(* IEC 61131-3 sources: deprecated-refusr-repo/samples (part 19) *)

(* ---- RND-EXPR_audio-kudos-nifty.st ---- *)
(*
This code implements a randomly grown symbolic expression:

IN3 | (xor(xor(IN43 | ((xor(xor(!(((xor(xor(IN13, IN9 | false), xor(xor(IN25, IN14), IN11))) | (xor(xor(xor(xor(IN36, IN12), IN39), IN13 & IN34), IN47))) | (xor(xor(IN5, (IN1 & IN27) | (!(IN46))), !(!(IN21))))), IN37), xor(xor(!(!(IN1)), !((xor(xor(IN30, false), xor(xor(IN49, IN30), IN25))) & (!(xor(xor(IN21, IN32), IN27))))), (xor(xor(!(xor(xor(IN12, IN39), IN41)), (IN22 & IN36) & (IN27 | IN16)), IN15)) | (!((IN24 | IN40) | (!(IN45))))))) & (xor(xor(!((!((false | IN41) & (!(IN49)))) | (((IN6 & IN32) & IN14) & (!(IN27 & IN33)))), xor(xor(xor(xor(IN38, (!(IN43 & IN26)) & ((IN34 & IN40) & (IN5 & IN12))), !(xor(xor(xor(xor(IN8, IN19), IN14), IN15 & IN11), IN30 & IN31))), ((xor(xor(IN24, IN1 | IN19), true | IN1)) & IN27) & ((IN25 | (IN21 | IN15)) & (IN13 & (IN19 & IN30)))), (((IN33 & true) | (IN35 | IN7)) & (xor(xor(true | IN16, IN48), IN43 & IN22))) & ((!(xor(xor(IN38, IN35), IN42))) & (!(IN39))))), xor(xor(IN6, (xor(xor(xor(xor(xor(xor(IN6, IN45), IN26), !(IN35)), IN32 | IN15), (!(IN15)) & (IN36 | IN34)), (xor(xor(IN47, IN47), IN44)) & (!(IN14)))) & (((IN13 & IN4) | (IN1 | IN38)) | ((IN46 & IN11) & (IN32 | IN24)))), IN18)))), !(xor(xor(!(!(xor(xor(IN1, !((xor(xor(IN33, IN25), IN4)) & (IN40 | IN38))), xor(xor(IN12, xor(xor(xor(xor(IN24, IN3), IN41), !(IN13)), IN50 & IN19)), (xor(xor(IN37, IN25), IN21)) | IN4)))), !(IN23)), (!((!((!(IN20)) & (IN23 & IN14))) | (IN43 | (xor(xor(IN27 & IN10, IN34), xor(xor(IN31, IN6), IN4)))))) | ((((!(IN27 | IN41)) | ((IN12 | IN28) | IN22)) & IN29) & (IN50 & (IN1 | ((xor(xor(IN49, IN28), IN4)) | (IN33 & IN4)))))))), (!((xor(xor((!(xor(xor(!(IN27), xor(xor(IN4, IN6), IN33)), IN31 & true))) | (!((xor(xor(IN40, IN39), IN27)) & (IN13 & IN12))), (((IN25 & IN4) & (!(IN17))) & (xor(xor(true | IN33, IN38), IN16))) & (xor(xor(IN44, !(xor(xor(IN27, IN40), IN11))), xor(xor(IN36 & IN37, IN15 | IN33), IN21)))), IN17 | (IN33 | ((IN2 & IN1) | IN33)))) & (((((IN33 & false) | (IN37 | IN18)) | (!(IN28))) & (xor(xor((IN38 | IN8) | (!(IN12)), !(IN1 | IN1)), IN30))) | (xor(xor((xor(xor(IN47 & IN24, IN47 & IN36), IN9)) & (!(IN31 & IN18)), xor(xor((!(IN49)) & IN4, (IN44 & IN19) | (IN26 | IN18)), !(!(IN34)))), !(IN32 & (IN33 | IN47))))))) | ((xor(xor(IN13, (!(true | (xor(xor(!(IN35), IN15 | IN4), xor(xor(IN35, IN27), IN15))))) & ((xor(xor(!(IN18 & IN31), IN22 | (IN7 & IN11)), !(xor(xor(IN37, IN45), IN24)))) & IN23)), IN35)) & IN5)))

*)

FUNCTION_BLOCK F_CollectInput
  VAR_IN_OUT
      Data : ARRAY[1..50] OF BOOL;
  END_VAR
  VAR_INPUT
      TICK  : BOOL := 0;
      IN1   : BOOL := 0;
      IN2   : BOOL := 0;
      IN3   : BOOL := 0;
      IN4   : BOOL := 0;
      IN5   : BOOL := 0;
      RESET : BOOL := FALSE;
  END_VAR
  VAR_OUTPUT
      Finished : BOOL;
  END_VAR
  VAR
      j    : USINT := 1;
      tock : BOOL  := 0;
  END_VAR
  IF NOT RESET AND tock = NOT TICK THEN
      Data[j]   := IN1;
      Data[j+1] := IN2;
      Data[j+2] := IN3;
      Data[j+3] := IN4;
      Data[j+4] := IN5;
      j := j + 5;
      tock := TICK;
  ELSE
      j := 1;
      tock := 0;
  END_IF;
  Finished := (j > 50);
END_FUNCTION_BLOCK

PROGRAM Boiler
  VAR
    Data  : ARRAY[1..50] OF BOOL;
    Ready : BOOL;
    CollectInput : F_CollectInput;
  END_VAR
  VAR
    TICK     AT %IX1.0 : BOOL;
    IN1      AT %IX0.3 : BOOL;
    IN2      AT %IX0.4 : BOOL;
    IN3      AT %IX0.5 : BOOL;
    IN4      AT %IX0.6 : BOOL;
    IN5      AT %IX0.7 : BOOL;
    OutReady AT %QX0.0 : BOOL := FALSE;
    FeedNext AT %QX0.1 : BOOL := FALSE;
    Out      AT %QX0.2 : BOOL;
  END_VAR
  CollectInput(TICK:=TICK, IN1:=IN1, IN2:=IN2, IN3:=IN3, IN4:=IN4, IN5:=IN5);
  Ready := CollectInput.Finished;
  FeedNext := 1;
  IF Ready THEN
    Out := (Data[3] OR (((Data[43] OR ((((NOT ((((Data[13] XOR (Data[9] OR FALSE)) XOR ((Data[25] XOR Data[14]) XOR Data[11])) OR ((((Data[36] XOR Data[12]) XOR Data[39]) XOR (Data[13] AND Data[34])) XOR Data[47])) OR ((Data[5] XOR ((Data[1] AND Data[27]) OR (NOT Data[46]))) XOR (NOT (NOT Data[21]))))) XOR Data[37]) XOR (((NOT (NOT Data[1])) XOR (NOT (((Data[30] XOR FALSE) XOR ((Data[49] XOR Data[30]) XOR Data[25])) AND (NOT ((Data[21] XOR Data[32]) XOR Data[27]))))) XOR ((((NOT ((Data[12] XOR Data[39]) XOR Data[41])) XOR ((Data[22] AND Data[36]) AND (Data[27] OR Data[16]))) XOR Data[15]) OR (NOT ((Data[24] OR Data[40]) OR (NOT Data[45])))))) AND (((NOT ((NOT ((FALSE OR Data[41]) AND (NOT Data[49]))) OR (((Data[6] AND Data[32]) AND Data[14]) AND (NOT (Data[27] AND Data[33]))))) XOR ((((Data[38] XOR ((NOT (Data[43] AND Data[26])) AND ((Data[34] AND Data[40]) AND (Data[5] AND Data[12])))) XOR (NOT ((((Data[8] XOR Data[19]) XOR Data[14]) XOR (Data[15] AND Data[11])) XOR (Data[30] AND Data[31])))) XOR ((((Data[24] XOR (Data[1] OR Data[19])) XOR (TRUE OR Data[1])) AND Data[27]) AND ((Data[25] OR (Data[21] OR Data[15])) AND (Data[13] AND (Data[19] AND Data[30]))))) XOR ((((Data[33] AND TRUE) OR (Data[35] OR Data[7])) AND (((TRUE OR Data[16]) XOR Data[48]) XOR (Data[43] AND Data[22]))) AND ((NOT ((Data[38] XOR Data[35]) XOR Data[42])) AND (NOT Data[39]))))) XOR ((Data[6] XOR (((((((Data[6] XOR Data[45]) XOR Data[26]) XOR (NOT Data[35])) XOR (Data[32] OR Data[15])) XOR ((NOT Data[15]) AND (Data[36] OR Data[34]))) XOR (((Data[47] XOR Data[47]) XOR Data[44]) AND (NOT Data[14]))) AND (((Data[13] AND Data[4]) OR (Data[1] OR Data[38])) OR ((Data[46] AND Data[11]) AND (Data[32] OR Data[24]))))) XOR Data[18])))) XOR (NOT (((NOT (NOT ((Data[1] XOR (NOT (((Data[33] XOR Data[25]) XOR Data[4]) AND (Data[40] OR Data[38])))) XOR ((Data[12] XOR ((((Data[24] XOR Data[3]) XOR Data[41]) XOR (NOT Data[13])) XOR (Data[50] AND Data[19]))) XOR (((Data[37] XOR Data[25]) XOR Data[21]) OR Data[4]))))) XOR (NOT Data[23])) XOR ((NOT ((NOT ((NOT Data[20]) AND (Data[23] AND Data[14]))) OR (Data[43] OR (((Data[27] AND Data[10]) XOR Data[34]) XOR ((Data[31] XOR Data[6]) XOR Data[4]))))) OR ((((NOT (Data[27] OR Data[41])) OR ((Data[12] OR Data[28]) OR Data[22])) AND Data[29]) AND (Data[50] AND (Data[1] OR (((Data[49] XOR Data[28]) XOR Data[4]) OR (Data[33] AND Data[4]))))))))) XOR ((NOT (((((NOT (((NOT Data[27]) XOR ((Data[4] XOR Data[6]) XOR Data[33])) XOR (Data[31] AND TRUE))) OR (NOT (((Data[40] XOR Data[39]) XOR Data[27]) AND (Data[13] AND Data[12])))) XOR ((((Data[25] AND Data[4]) AND (NOT Data[17])) AND (((TRUE OR Data[33]) XOR Data[38]) XOR Data[16])) AND ((Data[44] XOR (NOT ((Data[27] XOR Data[40]) XOR Data[11]))) XOR (((Data[36] AND Data[37]) XOR (Data[15] OR Data[33])) XOR Data[21])))) XOR (Data[17] OR (Data[33] OR ((Data[2] AND Data[1]) OR Data[33])))) AND (((((Data[33] AND FALSE) OR (Data[37] OR Data[18])) OR (NOT Data[28])) AND ((((Data[38] OR Data[8]) OR (NOT Data[12])) XOR (NOT (Data[1] OR Data[1]))) XOR Data[30])) OR ((((((Data[47] AND Data[24]) XOR (Data[47] AND Data[36])) XOR Data[9]) AND (NOT (Data[31] AND Data[18]))) XOR ((((NOT Data[49]) AND Data[4]) XOR ((Data[44] AND Data[19]) OR (Data[26] OR Data[18]))) XOR (NOT (NOT Data[34])))) XOR (NOT (Data[32] AND (Data[33] OR Data[47]))))))) OR (((Data[13] XOR ((NOT (TRUE OR (((NOT Data[35]) XOR (Data[15] OR Data[4])) XOR ((Data[35] XOR Data[27]) XOR Data[15])))) AND ((((NOT (Data[18] AND Data[31])) XOR (Data[22] OR (Data[7] AND Data[11]))) XOR (NOT ((Data[37] XOR Data[45]) XOR Data[24]))) AND Data[23]))) XOR Data[35]) AND Data[5]))));
    OutReady := 1;
    CollectInput(RESET:=TRUE);
  END_IF;
END_PROGRAM

CONFIGURATION Config0
  RESOURCE Res0 ON PLC
    TASK task0(INTERVAL := T#20ms,PRIORITY := 0);
    PROGRAM instance0 WITH task0 : Boiler;
  END_RESOURCE
END_CONFIGURATION

(* ---- RND-EXPR_awoke-fount-idled.st ---- *)
(*
This code implements a randomly grown symbolic expression:

!(xor(xor(IN7, (xor(xor(IN10 | (xor(xor(IN35 & (((xor(xor(IN23, IN37), IN21)) & (IN38 & IN15)) | (xor(xor(xor(xor(IN32, IN34), IN21), false & IN13), IN2 | IN26))), IN35 & (((xor(xor(IN7, IN2), false)) | (!(IN1))) | (xor(xor(!(IN25), xor(xor(IN45, IN1), IN42)), IN26 | IN16)))), xor(xor((xor(xor(!(IN35), IN47 | IN5), IN39 & IN10)) & ((xor(xor(IN16, IN37), IN23)) | (!(IN48))), !(IN46)), !(!(!(IN21)))))), IN28), false)) & (xor(xor(xor(xor((((xor(xor(xor(xor(IN46, IN37), IN44), IN29 & IN42), IN10 | false)) | (xor(xor(IN38 & false, IN30 & IN3), true))) | (((xor(xor(IN14, IN23), IN50)) & (xor(xor(IN24, IN27), IN22))) | ((xor(xor(IN18, IN21), IN34)) & (true | IN4)))) & (xor(xor((xor(xor(xor(xor(IN29, IN24), true), IN12 & IN14), IN2 | IN19)) & (!(IN30 & IN14)), (IN10 | (!(IN9))) | ((IN42 & IN44) & (IN33 & IN25))), IN5)), IN3 & ((xor(xor((IN36 & IN29) & (IN6 | IN45), xor(xor(!(IN2), !(IN10)), IN20)), IN43)) & (!((IN33 | IN35) | (xor(xor(IN50, IN35), IN48)))))), xor(xor((xor(xor(!(!(IN46)), IN34 | (IN35 | IN49)), (!(IN34)) & (IN10 & IN4))) & (IN15 | IN25), IN22), (xor(xor(xor(xor(IN30, IN12 | IN23), !(IN14)), IN1), (IN4 | IN32) & (!(IN48)))) | (((xor(xor(IN50, true), IN31)) & (xor(xor(IN22, IN32), IN34))) | (xor(xor(IN37, !(IN49)), IN22))))), xor(xor(!(xor(xor(xor(xor((IN48 & IN24) | (xor(xor(IN41, IN39), IN11)), IN14), IN11), IN39 & (!(IN10 | IN49))), IN44)), ((!(!(!(IN50)))) & ((xor(xor(IN35, !(IN50)), IN32 | IN49)) & (xor(xor(IN21 & IN42, true & IN25), IN4 & IN31)))) | (((!(IN21)) | (!(xor(xor(IN1, IN30), IN46)))) & (((IN6 | IN8) & (xor(xor(IN43, IN10), false))) | IN6))), xor(xor((xor(xor((IN34 | IN3) & (!(IN18)), (!(IN14)) & true), xor(xor(xor(xor(IN15, IN7), IN34), !(IN31)), IN20 | IN18))) | (((IN1 | IN1) & (IN5 | IN27)) | IN17), xor(xor((xor(xor(xor(xor(IN32, IN10), IN1), IN35 | IN32), IN8)) & (IN11 & (IN14 | IN16)), !((IN20 & IN44) | (IN6 | IN15))), (xor(xor(IN35 | IN40, !(IN35)), IN3 | IN48)) | (!(IN46)))), (!(IN14)) & IN7))), (xor(xor(!(xor(xor(IN18, xor(xor(IN24 & IN23, !(IN40)), xor(xor(IN27, IN31), IN35))), !(xor(xor(false, IN48), IN6)))), (!((IN23 | IN37) & (IN8 | IN41))) & IN25), IN5 | (((xor(xor(IN41, IN26), IN3)) & (IN46 | IN22)) | ((IN49 & IN45) & (IN42 & IN16))))) | ((((!(IN47)) | true) & (IN30 | ((IN46 & IN30) | (!(IN43))))) | (((xor(xor(IN37, !(IN40)), !(IN4))) | (IN11 & (!(IN40)))) | (xor(xor(xor(xor(IN46 | IN15, IN9 | IN2), !(IN15)), xor(xor(!(IN46), false), IN36 & IN44)), !(!(IN27))))))))), !(IN35 & (xor(xor((xor(xor(xor(xor(!(xor(xor(IN12, IN9), IN31)), (xor(xor(IN35, IN38), IN3)) | (xor(xor(IN47, IN13), IN8))), (IN36 & false) | (IN13 | IN46)), IN19), (IN47 & (IN46 | IN35)) | IN25)) & (xor(xor(xor(xor((IN14 | IN37) | (IN10 | IN3), IN39 & IN30), xor(xor(IN33 & IN5, xor(xor(IN39, IN48), IN16)), !(IN33))), !(IN38)), !(!(IN33 | IN3)))), IN48), IN20)))))

*)

FUNCTION_BLOCK F_CollectInput
  VAR_IN_OUT
      Data : ARRAY[1..50] OF BOOL;
  END_VAR
  VAR_INPUT
      TICK  : BOOL := 0;
      IN1   : BOOL := 0;
      IN2   : BOOL := 0;
      IN3   : BOOL := 0;
      IN4   : BOOL := 0;
      IN5   : BOOL := 0;
      RESET : BOOL := FALSE;
  END_VAR
  VAR_OUTPUT
      Finished : BOOL;
  END_VAR
  VAR
      j    : USINT := 1;
      tock : BOOL  := 0;
  END_VAR
  IF NOT RESET AND tock = NOT TICK THEN
      Data[j]   := IN1;
      Data[j+1] := IN2;
      Data[j+2] := IN3;
      Data[j+3] := IN4;
      Data[j+4] := IN5;
      j := j + 5;
      tock := TICK;
  ELSE
      j := 1;
      tock := 0;
  END_IF;
  Finished := (j > 50);
END_FUNCTION_BLOCK

PROGRAM Boiler
  VAR
    Data  : ARRAY[1..50] OF BOOL;
    Ready : BOOL;
    CollectInput : F_CollectInput;
  END_VAR
  VAR
    TICK     AT %IX1.0 : BOOL;
    IN1      AT %IX0.3 : BOOL;
    IN2      AT %IX0.4 : BOOL;
    IN3      AT %IX0.5 : BOOL;
    IN4      AT %IX0.6 : BOOL;
    IN5      AT %IX0.7 : BOOL;
    OutReady AT %QX0.0 : BOOL := FALSE;
    FeedNext AT %QX0.1 : BOOL := FALSE;
    Out      AT %QX0.2 : BOOL;
  END_VAR
  CollectInput(TICK:=TICK, IN1:=IN1, IN2:=IN2, IN3:=IN3, IN4:=IN4, IN5:=IN5);
  Ready := CollectInput.Finished;
  FeedNext := 1;
  IF Ready THEN
    Out := (NOT ((Data[7] XOR ((((Data[10] OR (((Data[35] AND ((((Data[23] XOR Data[37]) XOR Data[21]) AND (Data[38] AND Data[15])) OR ((((Data[32] XOR Data[34]) XOR Data[21]) XOR (FALSE AND Data[13])) XOR (Data[2] OR Data[26])))) XOR (Data[35] AND ((((Data[7] XOR Data[2]) XOR FALSE) OR (NOT Data[1])) OR (((NOT Data[25]) XOR ((Data[45] XOR Data[1]) XOR Data[42])) XOR (Data[26] OR Data[16]))))) XOR ((((((NOT Data[35]) XOR (Data[47] OR Data[5])) XOR (Data[39] AND Data[10])) AND (((Data[16] XOR Data[37]) XOR Data[23]) OR (NOT Data[48]))) XOR (NOT Data[46])) XOR (NOT (NOT (NOT Data[21])))))) XOR Data[28]) XOR FALSE) AND (((((((((((Data[46] XOR Data[37]) XOR Data[44]) XOR (Data[29] AND Data[42])) XOR (Data[10] OR FALSE)) OR (((Data[38] AND FALSE) XOR (Data[30] AND Data[3])) XOR TRUE)) OR ((((Data[14] XOR Data[23]) XOR Data[50]) AND ((Data[24] XOR Data[27]) XOR Data[22])) OR (((Data[18] XOR Data[21]) XOR Data[34]) AND (TRUE OR Data[4])))) AND (((((((Data[29] XOR Data[24]) XOR TRUE) XOR (Data[12] AND Data[14])) XOR (Data[2] OR Data[19])) AND (NOT (Data[30] AND Data[14]))) XOR ((Data[10] OR (NOT Data[9])) OR ((Data[42] AND Data[44]) AND (Data[33] AND Data[25])))) XOR Data[5])) XOR (Data[3] AND (((((Data[36] AND Data[29]) AND (Data[6] OR Data[45])) XOR (((NOT Data[2]) XOR (NOT Data[10])) XOR Data[20])) XOR Data[43]) AND (NOT ((Data[33] OR Data[35]) OR ((Data[50] XOR Data[35]) XOR Data[48])))))) XOR ((((((NOT (NOT Data[46])) XOR (Data[34] OR (Data[35] OR Data[49]))) XOR ((NOT Data[34]) AND (Data[10] AND Data[4]))) AND (Data[15] OR Data[25])) XOR Data[22]) XOR (((((Data[30] XOR (Data[12] OR Data[23])) XOR (NOT Data[14])) XOR Data[1]) XOR ((Data[4] OR Data[32]) AND (NOT Data[48]))) OR ((((Data[50] XOR TRUE) XOR Data[31]) AND ((Data[22] XOR Data[32]) XOR Data[34])) OR ((Data[37] XOR (NOT Data[49])) XOR Data[22]))))) XOR (((NOT ((((((Data[48] AND Data[24]) OR ((Data[41] XOR Data[39]) XOR Data[11])) XOR Data[14]) XOR Data[11]) XOR (Data[39] AND (NOT (Data[10] OR Data[49])))) XOR Data[44])) XOR (((NOT (NOT (NOT Data[50]))) AND (((Data[35] XOR (NOT Data[50])) XOR (Data[32] OR Data[49])) AND (((Data[21] AND Data[42]) XOR (TRUE AND Data[25])) XOR (Data[4] AND Data[31])))) OR (((NOT Data[21]) OR (NOT ((Data[1] XOR Data[30]) XOR Data[46]))) AND (((Data[6] OR Data[8]) AND ((Data[43] XOR Data[10]) XOR FALSE)) OR Data[6])))) XOR (((((((Data[34] OR Data[3]) AND (NOT Data[18])) XOR ((NOT Data[14]) AND TRUE)) XOR ((((Data[15] XOR Data[7]) XOR Data[34]) XOR (NOT Data[31])) XOR (Data[20] OR Data[18]))) OR (((Data[1] OR Data[1]) AND (Data[5] OR Data[27])) OR Data[17])) XOR (((((((Data[32] XOR Data[10]) XOR Data[1]) XOR (Data[35] OR Data[32])) XOR Data[8]) AND (Data[11] AND (Data[14] OR Data[16]))) XOR (NOT ((Data[20] AND Data[44]) OR (Data[6] OR Data[15])))) XOR ((((Data[35] OR Data[40]) XOR (NOT Data[35])) XOR (Data[3] OR Data[48])) OR (NOT Data[46])))) XOR ((NOT Data[14]) AND Data[7])))) XOR ((((NOT ((Data[18] XOR (((Data[24] AND Data[23]) XOR (NOT Data[40])) XOR ((Data[27] XOR Data[31]) XOR Data[35]))) XOR (NOT ((FALSE XOR Data[48]) XOR Data[6])))) XOR ((NOT ((Data[23] OR Data[37]) AND (Data[8] OR Data[41]))) AND Data[25])) XOR (Data[5] OR ((((Data[41] XOR Data[26]) XOR Data[3]) AND (Data[46] OR Data[22])) OR ((Data[49] AND Data[45]) AND (Data[42] AND Data[16]))))) OR ((((NOT Data[47]) OR TRUE) AND (Data[30] OR ((Data[46] AND Data[30]) OR (NOT Data[43])))) OR ((((Data[37] XOR (NOT Data[40])) XOR (NOT Data[4])) OR (Data[11] AND (NOT Data[40]))) OR (((((Data[46] OR Data[15]) XOR (Data[9] OR Data[2])) XOR (NOT Data[15])) XOR (((NOT Data[46]) XOR FALSE) XOR (Data[36] AND Data[44]))) XOR (NOT (NOT Data[27]))))))))) XOR (NOT (Data[35] AND ((((((((NOT ((Data[12] XOR Data[9]) XOR Data[31])) XOR (((Data[35] XOR Data[38]) XOR Data[3]) OR ((Data[47] XOR Data[13]) XOR Data[8]))) XOR ((Data[36] AND FALSE) OR (Data[13] OR Data[46]))) XOR Data[19]) XOR ((Data[47] AND (Data[46] OR Data[35])) OR Data[25])) AND ((((((Data[14] OR Data[37]) OR (Data[10] OR Data[3])) XOR (Data[39] AND Data[30])) XOR (((Data[33] AND Data[5]) XOR ((Data[39] XOR Data[48]) XOR Data[16])) XOR (NOT Data[33]))) XOR (NOT Data[38])) XOR (NOT (NOT (Data[33] OR Data[3]))))) XOR Data[48]) XOR Data[20])))));
    OutReady := 1;
    CollectInput(RESET:=TRUE);
  END_IF;
END_PROGRAM

CONFIGURATION Config0
  RESOURCE Res0 ON PLC
    TASK task0(INTERVAL := T#20ms,PRIORITY := 0);
    PROGRAM instance0 WITH task0 : Boiler;
  END_RESOURCE
END_CONFIGURATION

(* ---- RND-EXPR_balmy-flubs-lives.st ---- *)
(*
This code implements a randomly grown symbolic expression:

(!(IN49)) & IN46

*)

FUNCTION_BLOCK F_CollectInput
  VAR_IN_OUT
      Data : ARRAY[1..50] OF BOOL;
  END_VAR
  VAR_INPUT
      TICK  : BOOL := 0;
      IN1   : BOOL := 0;
      IN2   : BOOL := 0;
      IN3   : BOOL := 0;
      IN4   : BOOL := 0;
      IN5   : BOOL := 0;
      RESET : BOOL := FALSE;
  END_VAR
  VAR_OUTPUT
      Finished : BOOL;
  END_VAR
  VAR
      j    : USINT := 1;
      tock : BOOL  := 0;
  END_VAR
  IF NOT RESET AND tock = NOT TICK THEN
      Data[j]   := IN1;
      Data[j+1] := IN2;
      Data[j+2] := IN3;
      Data[j+3] := IN4;
      Data[j+4] := IN5;
      j := j + 5;
      tock := TICK;
  ELSE
      j := 1;
      tock := 0;
  END_IF;
  Finished := (j > 50);
END_FUNCTION_BLOCK

PROGRAM Boiler
  VAR
    Data  : ARRAY[1..50] OF BOOL;
    Ready : BOOL;
    CollectInput : F_CollectInput;
  END_VAR
  VAR
    TICK     AT %IX1.0 : BOOL;
    IN1      AT %IX0.3 : BOOL;
    IN2      AT %IX0.4 : BOOL;
    IN3      AT %IX0.5 : BOOL;
    IN4      AT %IX0.6 : BOOL;
    IN5      AT %IX0.7 : BOOL;
    OutReady AT %QX0.0 : BOOL := FALSE;
    FeedNext AT %QX0.1 : BOOL := FALSE;
    Out      AT %QX0.2 : BOOL;
  END_VAR
  CollectInput(TICK:=TICK, IN1:=IN1, IN2:=IN2, IN3:=IN3, IN4:=IN4, IN5:=IN5);
  Ready := CollectInput.Finished;
  FeedNext := 1;
  IF Ready THEN
    Out := ((NOT Data[49]) AND Data[46]);
    OutReady := 1;
    CollectInput(RESET:=TRUE);
  END_IF;
END_PROGRAM

CONFIGURATION Config0
  RESOURCE Res0 ON PLC
    TASK task0(INTERVAL := T#20ms,PRIORITY := 0);
    PROGRAM instance0 WITH task0 : Boiler;
  END_RESOURCE
END_CONFIGURATION

(* ---- RND-EXPR_baton-smear-tarot.st ---- *)
(*
This code implements a randomly grown symbolic expression:

xor(xor(!((((IN19 | ((!(xor(xor(IN42 | IN9, IN18), IN43))) & (IN45 & (!(xor(xor(IN20, IN7), IN15)))))) | (xor(xor(IN2, (((xor(xor(IN43, IN1), IN41)) | (xor(xor(IN13, IN45), IN31))) & ((IN14 & IN3) | (IN11 | IN19))) | IN16), IN5 | IN40))) & IN38) & (IN44 | (IN29 & IN45))), xor(xor(IN21, IN35 & (!(IN21))), (!(xor(xor(xor(xor((!(IN16 | (xor(xor(IN8, IN25), IN37)))) & IN21, IN12), (!((IN32 & IN11) & (IN26 | IN3))) | (xor(xor(xor(xor(IN18 | IN31, IN48 | IN23), IN26 & IN42), !(IN24)), (IN22 & IN13) & (IN25 | IN12)))), IN16), IN13))) | (((!((((IN13 & IN39) & (!(IN34))) | IN2) | (!(!(xor(xor(IN23, IN32), IN28)))))) | (xor(xor(xor(xor((xor(xor(IN38 & IN21, IN45 | IN35), IN21 & IN26)) | IN1, ((IN23 | IN23) | IN17) & (!(IN20 & IN9))), IN39), !(!(xor(xor(IN26 & IN43, IN40 & IN33), false | IN33)))), IN49))) | IN3))), (!(!(!(IN2 & IN26)))) & (xor(xor((xor(xor((xor(xor(IN27, xor(xor(IN42 & (!(IN35)), (IN3 | IN32) & (IN4 | IN35)), (!(IN32)) & IN47)), (xor(xor(xor(xor(IN13, IN2), IN28), IN9 | IN42), !(IN30))) | ((IN9 | IN14) & (IN44 & IN28)))) & (!(IN21 | ((IN1 | IN41) & (IN6 | IN3)))), !(((!(IN41)) | IN41) & (IN13 | ((IN13 & IN10) & (xor(xor(IN27, IN13), IN7)))))), !(xor(xor(IN18, IN9), (!(IN38 & IN26)) & (xor(xor(IN21 | IN41, xor(xor(IN23, IN37), IN28)), !(IN7))))))) & ((!(xor(xor((IN17 & (!(IN29))) & ((IN22 & IN31) | (xor(xor(IN13, IN47), IN2))), ((!(IN7)) | IN4) | (xor(xor(!(IN19), !(IN19)), IN31))), !((xor(xor(IN8, IN12), false)) & (IN25 | IN21))))) & (IN5 | (xor(xor(xor(xor(xor(xor(xor(xor(IN14, IN16), IN50), IN9), IN44), xor(xor(xor(xor(IN19, IN1), IN13), IN2 & IN36), IN40)), !(IN10 | IN39)), IN20), (IN4 & (!(IN21))) & (IN8 | (IN30 & IN12)))))), (xor(xor((!((xor(xor(IN50 | IN6, IN28 & IN9), IN23)) | (xor(xor(IN41 | IN44, IN7 | IN29), !(IN26))))) | (((xor(xor(IN4, IN43 | IN10), IN17 & IN40)) & ((IN49 & IN39) & (xor(xor(IN18, IN39), IN12)))) & (!(IN11 & (IN26 | IN30)))), IN13), IN2 | ((((xor(xor(IN32, IN41), IN4)) & IN43) & ((IN18 | IN10) | (xor(xor(IN22, IN16), IN42)))) & (IN22 | (xor(xor(IN18 & IN35, IN14), IN20 & IN8)))))) & (((xor(xor(((IN6 & IN44) | (xor(xor(IN11, IN45), true))) | IN11, true), xor(xor((xor(xor(IN8, true), IN25)) & (xor(xor(IN39, IN32), IN11)), !(IN21 | IN28)), IN6))) | ((xor(xor(IN14, (!(IN16)) & (!(IN29))), xor(xor(IN27 | IN23, IN13), xor(xor(IN12, IN25), IN31)))) | (xor(xor(xor(xor(IN11 | IN50, !(IN48)), !(IN48)), IN14), IN27)))) | (!(IN34 & (((IN3 | IN14) | (true & IN17)) & ((xor(xor(IN39, IN50), IN5)) | (IN4 | IN18))))))), IN5)))

*)

FUNCTION_BLOCK F_CollectInput
  VAR_IN_OUT
      Data : ARRAY[1..50] OF BOOL;
  END_VAR
  VAR_INPUT
      TICK  : BOOL := 0;
      IN1   : BOOL := 0;
      IN2   : BOOL := 0;
      IN3   : BOOL := 0;
      IN4   : BOOL := 0;
      IN5   : BOOL := 0;
      RESET : BOOL := FALSE;
  END_VAR
  VAR_OUTPUT
      Finished : BOOL;
  END_VAR
  VAR
      j    : USINT := 1;
      tock : BOOL  := 0;
  END_VAR
  IF NOT RESET AND tock = NOT TICK THEN
      Data[j]   := IN1;
      Data[j+1] := IN2;
      Data[j+2] := IN3;
      Data[j+3] := IN4;
      Data[j+4] := IN5;
      j := j + 5;
      tock := TICK;
  ELSE
      j := 1;
      tock := 0;
  END_IF;
  Finished := (j > 50);
END_FUNCTION_BLOCK

PROGRAM Boiler
  VAR
    Data  : ARRAY[1..50] OF BOOL;
    Ready : BOOL;
    CollectInput : F_CollectInput;
  END_VAR
  VAR
    TICK     AT %IX1.0 : BOOL;
    IN1      AT %IX0.3 : BOOL;
    IN2      AT %IX0.4 : BOOL;
    IN3      AT %IX0.5 : BOOL;
    IN4      AT %IX0.6 : BOOL;
    IN5      AT %IX0.7 : BOOL;
    OutReady AT %QX0.0 : BOOL := FALSE;
    FeedNext AT %QX0.1 : BOOL := FALSE;
    Out      AT %QX0.2 : BOOL;
  END_VAR
  CollectInput(TICK:=TICK, IN1:=IN1, IN2:=IN2, IN3:=IN3, IN4:=IN4, IN5:=IN5);
  Ready := CollectInput.Finished;
  FeedNext := 1;
  IF Ready THEN
    Out := (((NOT ((((Data[19] OR ((NOT (((Data[42] OR Data[9]) XOR Data[18]) XOR Data[43])) AND (Data[45] AND (NOT ((Data[20] XOR Data[7]) XOR Data[15]))))) OR ((Data[2] XOR (((((Data[43] XOR Data[1]) XOR Data[41]) OR ((Data[13] XOR Data[45]) XOR Data[31])) AND ((Data[14] AND Data[3]) OR (Data[11] OR Data[19]))) OR Data[16])) XOR (Data[5] OR Data[40]))) AND Data[38]) AND (Data[44] OR (Data[29] AND Data[45])))) XOR ((Data[21] XOR (Data[35] AND (NOT Data[21]))) XOR ((NOT ((((((NOT (Data[16] OR ((Data[8] XOR Data[25]) XOR Data[37]))) AND Data[21]) XOR Data[12]) XOR ((NOT ((Data[32] AND Data[11]) AND (Data[26] OR Data[3]))) OR (((((Data[18] OR Data[31]) XOR (Data[48] OR Data[23])) XOR (Data[26] AND Data[42])) XOR (NOT Data[24])) XOR ((Data[22] AND Data[13]) AND (Data[25] OR Data[12]))))) XOR Data[16]) XOR Data[13])) OR (((NOT ((((Data[13] AND Data[39]) AND (NOT Data[34])) OR Data[2]) OR (NOT (NOT ((Data[23] XOR Data[32]) XOR Data[28]))))) OR ((((((((Data[38] AND Data[21]) XOR (Data[45] OR Data[35])) XOR (Data[21] AND Data[26])) OR Data[1]) XOR (((Data[23] OR Data[23]) OR Data[17]) AND (NOT (Data[20] AND Data[9])))) XOR Data[39]) XOR (NOT (NOT (((Data[26] AND Data[43]) XOR (Data[40] AND Data[33])) XOR (FALSE OR Data[33]))))) XOR Data[49])) OR Data[3])))) XOR ((NOT (NOT (NOT (Data[2] AND Data[26])))) AND ((((((((Data[27] XOR (((Data[42] AND (NOT Data[35])) XOR ((Data[3] OR Data[32]) AND (Data[4] OR Data[35]))) XOR ((NOT Data[32]) AND Data[47]))) XOR (((((Data[13] XOR Data[2]) XOR Data[28]) XOR (Data[9] OR Data[42])) XOR (NOT Data[30])) OR ((Data[9] OR Data[14]) AND (Data[44] AND Data[28])))) AND (NOT (Data[21] OR ((Data[1] OR Data[41]) AND (Data[6] OR Data[3]))))) XOR (NOT (((NOT Data[41]) OR Data[41]) AND (Data[13] OR ((Data[13] AND Data[10]) AND ((Data[27] XOR Data[13]) XOR Data[7])))))) XOR (NOT ((Data[18] XOR Data[9]) XOR ((NOT (Data[38] AND Data[26])) AND (((Data[21] OR Data[41]) XOR ((Data[23] XOR Data[37]) XOR Data[28])) XOR (NOT Data[7])))))) AND ((NOT ((((Data[17] AND (NOT Data[29])) AND ((Data[22] AND Data[31]) OR ((Data[13] XOR Data[47]) XOR Data[2]))) XOR (((NOT Data[7]) OR Data[4]) OR (((NOT Data[19]) XOR (NOT Data[19])) XOR Data[31]))) XOR (NOT (((Data[8] XOR Data[12]) XOR FALSE) AND (Data[25] OR Data[21]))))) AND (Data[5] OR ((((((((Data[14] XOR Data[16]) XOR Data[50]) XOR Data[9]) XOR Data[44]) XOR ((((Data[19] XOR Data[1]) XOR Data[13]) XOR (Data[2] AND Data[36])) XOR Data[40])) XOR (NOT (Data[10] OR Data[39]))) XOR Data[20]) XOR ((Data[4] AND (NOT Data[21])) AND (Data[8] OR (Data[30] AND Data[12]))))))) XOR (((((NOT ((((Data[50] OR Data[6]) XOR (Data[28] AND Data[9])) XOR Data[23]) OR (((Data[41] OR Data[44]) XOR (Data[7] OR Data[29])) XOR (NOT Data[26])))) OR ((((Data[4] XOR (Data[43] OR Data[10])) XOR (Data[17] AND Data[40])) AND ((Data[49] AND Data[39]) AND ((Data[18] XOR Data[39]) XOR Data[12]))) AND (NOT (Data[11] AND (Data[26] OR Data[30]))))) XOR Data[13]) XOR (Data[2] OR (((((Data[32] XOR Data[41]) XOR Data[4]) AND Data[43]) AND ((Data[18] OR Data[10]) OR ((Data[22] XOR Data[16]) XOR Data[42]))) AND (Data[22] OR (((Data[18] AND Data[35]) XOR Data[14]) XOR (Data[20] AND Data[8])))))) AND (((((((Data[6] AND Data[44]) OR ((Data[11] XOR Data[45]) XOR TRUE)) OR Data[11]) XOR TRUE) XOR (((((Data[8] XOR TRUE) XOR Data[25]) AND ((Data[39] XOR Data[32]) XOR Data[11])) XOR (NOT (Data[21] OR Data[28]))) XOR Data[6])) OR (((Data[14] XOR ((NOT Data[16]) AND (NOT Data[29]))) XOR (((Data[27] OR Data[23]) XOR Data[13]) XOR ((Data[12] XOR Data[25]) XOR Data[31]))) OR (((((Data[11] OR Data[50]) XOR (NOT Data[48])) XOR (NOT Data[48])) XOR Data[14]) XOR Data[27]))) OR (NOT (Data[34] AND (((Data[3] OR Data[14]) OR (TRUE AND Data[17])) AND (((Data[39] XOR Data[50]) XOR Data[5]) OR (Data[4] OR Data[18])))))))) XOR Data[5])));
    OutReady := 1;
    CollectInput(RESET:=TRUE);
  END_IF;
END_PROGRAM

CONFIGURATION Config0
  RESOURCE Res0 ON PLC
    TASK task0(INTERVAL := T#20ms,PRIORITY := 0);
    PROGRAM instance0 WITH task0 : Boiler;
  END_RESOURCE
END_CONFIGURATION

(* ---- RND-EXPR_beads-fetal-heads.st ---- *)
(*
This code implements a randomly grown symbolic expression:

(((!((((!((IN5 & IN33) | (IN35 | IN14))) & (!(xor(xor(xor(xor(IN9, IN33), IN3), IN49 | IN12), IN43)))) & (IN16 | IN22)) | (IN9 | ((!(!(IN6 | IN26))) | (xor(xor(!(IN23 & true), (IN16 & IN22) | (!(IN20))), IN12)))))) | ((((xor(xor(xor(xor(IN28, (xor(xor(IN2, IN16), IN38)) & (xor(xor(IN24, IN21), IN24))), !(!(IN35))), !(IN31 & IN50)), xor(xor(xor(xor(!(IN26), xor(xor(IN1, IN45), IN39)), xor(xor(IN37, IN8), IN27)), xor(xor(IN1 | IN20, true & IN23), !(IN22))), xor(xor(!(IN39), xor(xor(IN1, IN47), IN27)), IN22 | IN16)))) | ((((!(IN26)) & (IN33 & IN22)) | ((xor(xor(IN45, IN43), IN41)) | (xor(xor(IN40, IN11), IN48)))) & ((xor(xor(IN24 | IN1, xor(xor(false, IN2), IN3)), IN5 | IN44)) | ((IN50 & IN2) | (!(IN49)))))) & (!(IN35))) | (xor(xor(!(!(!((IN50 | IN15) | (IN40 & IN2)))), ((((IN34 & IN30) | (IN45 | IN41)) & ((IN3 | IN38) | IN2)) & ((IN18 | (!(IN19))) | ((IN48 | IN30) & (!(IN7))))) | (!((xor(xor(IN29 | IN29, IN46 & IN22), IN18 | IN11)) & (!(IN49 & IN15))))), (!(xor(xor((!(IN26)) & IN35, (!(IN27)) & (IN23 | IN41)), IN49 | (!(IN47))))) & (!(!(xor(xor(xor(xor(IN8, IN50), IN23), xor(xor(IN6, IN18), IN22)), IN12 | IN7)))))))) & (xor(xor((((((!(xor(xor(IN14, IN6), IN3))) & IN4) | (!((IN14 & IN24) & (xor(xor(IN3, IN21), IN20))))) | ((((!(IN36)) & IN28) | IN2) & IN40)) | (!((IN13 | IN14) | (xor(xor((xor(xor(IN17, IN22), IN30)) & (IN35 | IN35), !(xor(xor(IN46, IN8), true))), !(IN22)))))) | (((!(IN50)) & (xor(xor(((xor(xor(IN26, IN26), IN31)) | (xor(xor(true, IN46), IN46))) | ((IN7 & IN17) & (xor(xor(IN5, IN38), IN21))), !((IN13 | IN22) & (IN16 | IN46))), xor(xor(xor(xor(IN37, IN36), xor(xor(IN2, IN44), IN18)), (IN28 & IN19) & (IN37 | IN20)), (IN24 & IN34) & (IN43 & IN45))))) | (IN39 | (((!(IN12)) | (IN21 | (!(IN38)))) & ((xor(xor(!(IN28), IN35 & IN29), !(IN50))) & ((xor(xor(IN42, IN19), IN47)) | IN42))))), xor(xor(!(xor(xor((((IN45 & IN48) & (xor(xor(IN21, IN32), IN36))) | ((IN20 | IN25) | (!(IN44)))) | (((!(IN28)) & IN15) | ((!(IN43)) | IN44)), xor(xor(xor(xor(IN7 | (xor(xor(IN43, IN3), IN10)), (!(IN1)) & IN48), !(xor(xor(IN34, IN19), IN42))), xor(xor((!(IN46)) | (IN32 & IN3), xor(xor(IN6 | IN20, !(IN29)), false & IN14)), !(!(IN20)))), xor(xor((xor(xor(IN24, IN27), IN37)) & IN26, !(IN33 & IN46)), !(xor(xor(IN7, IN41), IN38))))), xor(xor(!(!(IN26)), IN50), ((IN28 & IN17) & (xor(xor(IN4, IN38), IN9))) | ((IN16 | IN31) & (!(IN32)))))), !((!(!(!(xor(xor(IN9, IN1), IN39))))) & (!(IN1 & (!(xor(xor(IN20, IN38), false))))))), IN17)), xor(xor(xor(xor(((!(IN16 & (IN49 & IN24))) | (xor(xor((xor(xor(IN27, IN22), IN3)) | (xor(xor(false, IN46), IN40)), !(xor(xor(IN42, IN4), IN32))), IN22 & (xor(xor(IN8, IN30), IN3))))) | ((xor(xor(IN27 | (IN38 & IN36), xor(xor(IN24 | IN12, IN1 & IN37), !(IN39))), !(IN50 & IN47))) & (!((xor(xor(IN16, IN8), IN26)) | (IN49 | IN40)))), xor(xor(!(xor(xor(true, xor(xor(true, IN47), IN5 & IN29)), xor(xor(IN7 & IN8, IN19), !(IN23)))), (!(!(!(IN6)))) & IN9), true)), IN29), IN48), IN2)))) | IN11

*)

FUNCTION_BLOCK F_CollectInput
  VAR_IN_OUT
      Data : ARRAY[1..50] OF BOOL;
  END_VAR
  VAR_INPUT
      TICK  : BOOL := 0;
      IN1   : BOOL := 0;
      IN2   : BOOL := 0;
      IN3   : BOOL := 0;
      IN4   : BOOL := 0;
      IN5   : BOOL := 0;
      RESET : BOOL := FALSE;
  END_VAR
  VAR_OUTPUT
      Finished : BOOL;
  END_VAR
  VAR
      j    : USINT := 1;
      tock : BOOL  := 0;
  END_VAR
  IF NOT RESET AND tock = NOT TICK THEN
      Data[j]   := IN1;
      Data[j+1] := IN2;
      Data[j+2] := IN3;
      Data[j+3] := IN4;
      Data[j+4] := IN5;
      j := j + 5;
      tock := TICK;
  ELSE
      j := 1;
      tock := 0;
  END_IF;
  Finished := (j > 50);
END_FUNCTION_BLOCK

PROGRAM Boiler
  VAR
    Data  : ARRAY[1..50] OF BOOL;
    Ready : BOOL;
    CollectInput : F_CollectInput;
  END_VAR
  VAR
    TICK     AT %IX1.0 : BOOL;
    IN1      AT %IX0.3 : BOOL;
    IN2      AT %IX0.4 : BOOL;
    IN3      AT %IX0.5 : BOOL;
    IN4      AT %IX0.6 : BOOL;
    IN5      AT %IX0.7 : BOOL;
    OutReady AT %QX0.0 : BOOL := FALSE;
    FeedNext AT %QX0.1 : BOOL := FALSE;
    Out      AT %QX0.2 : BOOL;
  END_VAR
  CollectInput(TICK:=TICK, IN1:=IN1, IN2:=IN2, IN3:=IN3, IN4:=IN4, IN5:=IN5);
  Ready := CollectInput.Finished;
  FeedNext := 1;
  IF Ready THEN
    Out := ((((NOT ((((NOT ((Data[5] AND Data[33]) OR (Data[35] OR Data[14]))) AND (NOT ((((Data[9] XOR Data[33]) XOR Data[3]) XOR (Data[49] OR Data[12])) XOR Data[43]))) AND (Data[16] OR Data[22])) OR (Data[9] OR ((NOT (NOT (Data[6] OR Data[26]))) OR (((NOT (Data[23] AND TRUE)) XOR ((Data[16] AND Data[22]) OR (NOT Data[20]))) XOR Data[12]))))) OR (((((((Data[28] XOR (((Data[2] XOR Data[16]) XOR Data[38]) AND ((Data[24] XOR Data[21]) XOR Data[24]))) XOR (NOT (NOT Data[35]))) XOR (NOT (Data[31] AND Data[50]))) XOR (((((NOT Data[26]) XOR ((Data[1] XOR Data[45]) XOR Data[39])) XOR ((Data[37] XOR Data[8]) XOR Data[27])) XOR (((Data[1] OR Data[20]) XOR (TRUE AND Data[23])) XOR (NOT Data[22]))) XOR (((NOT Data[39]) XOR ((Data[1] XOR Data[47]) XOR Data[27])) XOR (Data[22] OR Data[16])))) OR ((((NOT Data[26]) AND (Data[33] AND Data[22])) OR (((Data[45] XOR Data[43]) XOR Data[41]) OR ((Data[40] XOR Data[11]) XOR Data[48]))) AND ((((Data[24] OR Data[1]) XOR ((FALSE XOR Data[2]) XOR Data[3])) XOR (Data[5] OR Data[44])) OR ((Data[50] AND Data[2]) OR (NOT Data[49]))))) AND (NOT Data[35])) OR (((NOT (NOT (NOT ((Data[50] OR Data[15]) OR (Data[40] AND Data[2]))))) XOR (((((Data[34] AND Data[30]) OR (Data[45] OR Data[41])) AND ((Data[3] OR Data[38]) OR Data[2])) AND ((Data[18] OR (NOT Data[19])) OR ((Data[48] OR Data[30]) AND (NOT Data[7])))) OR (NOT ((((Data[29] OR Data[29]) XOR (Data[46] AND Data[22])) XOR (Data[18] OR Data[11])) AND (NOT (Data[49] AND Data[15])))))) XOR ((NOT ((((NOT Data[26]) AND Data[35]) XOR ((NOT Data[27]) AND (Data[23] OR Data[41]))) XOR (Data[49] OR (NOT Data[47])))) AND (NOT (NOT ((((Data[8] XOR Data[50]) XOR Data[23]) XOR ((Data[6] XOR Data[18]) XOR Data[22])) XOR (Data[12] OR Data[7])))))))) AND ((((((((NOT ((Data[14] XOR Data[6]) XOR Data[3])) AND Data[4]) OR (NOT ((Data[14] AND Data[24]) AND ((Data[3] XOR Data[21]) XOR Data[20])))) OR ((((NOT Data[36]) AND Data[28]) OR Data[2]) AND Data[40])) OR (NOT ((Data[13] OR Data[14]) OR (((((Data[17] XOR Data[22]) XOR Data[30]) AND (Data[35] OR Data[35])) XOR (NOT ((Data[46] XOR Data[8]) XOR TRUE))) XOR (NOT Data[22]))))) OR (((NOT Data[50]) AND ((((((Data[26] XOR Data[26]) XOR Data[31]) OR ((TRUE XOR Data[46]) XOR Data[46])) OR ((Data[7] AND Data[17]) AND ((Data[5] XOR Data[38]) XOR Data[21]))) XOR (NOT ((Data[13] OR Data[22]) AND (Data[16] OR Data[46])))) XOR ((((Data[37] XOR Data[36]) XOR ((Data[2] XOR Data[44]) XOR Data[18])) XOR ((Data[28] AND Data[19]) AND (Data[37] OR Data[20]))) XOR ((Data[24] AND Data[34]) AND (Data[43] AND Data[45]))))) OR (Data[39] OR (((NOT Data[12]) OR (Data[21] OR (NOT Data[38]))) AND ((((NOT Data[28]) XOR (Data[35] AND Data[29])) XOR (NOT Data[50])) AND (((Data[42] XOR Data[19]) XOR Data[47]) OR Data[42])))))) XOR (((NOT ((((((Data[45] AND Data[48]) AND ((Data[21] XOR Data[32]) XOR Data[36])) OR ((Data[20] OR Data[25]) OR (NOT Data[44]))) OR (((NOT Data[28]) AND Data[15]) OR ((NOT Data[43]) OR Data[44]))) XOR (((((Data[7] OR ((Data[43] XOR Data[3]) XOR Data[10])) XOR ((NOT Data[1]) AND Data[48])) XOR (NOT ((Data[34] XOR Data[19]) XOR Data[42]))) XOR ((((NOT Data[46]) OR (Data[32] AND Data[3])) XOR (((Data[6] OR Data[20]) XOR (NOT Data[29])) XOR (FALSE AND Data[14]))) XOR (NOT (NOT Data[20])))) XOR (((((Data[24] XOR Data[27]) XOR Data[37]) AND Data[26]) XOR (NOT (Data[33] AND Data[46]))) XOR (NOT ((Data[7] XOR Data[41]) XOR Data[38]))))) XOR (((NOT (NOT Data[26])) XOR Data[50]) XOR (((Data[28] AND Data[17]) AND ((Data[4] XOR Data[38]) XOR Data[9])) OR ((Data[16] OR Data[31]) AND (NOT Data[32])))))) XOR (NOT ((NOT (NOT (NOT ((Data[9] XOR Data[1]) XOR Data[39])))) AND (NOT (Data[1] AND (NOT ((Data[20] XOR Data[38]) XOR FALSE))))))) XOR Data[17])) XOR (((((((NOT (Data[16] AND (Data[49] AND Data[24]))) OR (((((Data[27] XOR Data[22]) XOR Data[3]) OR ((FALSE XOR Data[46]) XOR Data[40])) XOR (NOT ((Data[42] XOR Data[4]) XOR Data[32]))) XOR (Data[22] AND ((Data[8] XOR Data[30]) XOR Data[3])))) OR ((((Data[27] OR (Data[38] AND Data[36])) XOR (((Data[24] OR Data[12]) XOR (Data[1] AND Data[37])) XOR (NOT Data[39]))) XOR (NOT (Data[50] AND Data[47]))) AND (NOT (((Data[16] XOR Data[8]) XOR Data[26]) OR (Data[49] OR Data[40]))))) XOR (((NOT ((TRUE XOR ((TRUE XOR Data[47]) XOR (Data[5] AND Data[29]))) XOR (((Data[7] AND Data[8]) XOR Data[19]) XOR (NOT Data[23])))) XOR ((NOT (NOT (NOT Data[6]))) AND Data[9])) XOR TRUE)) XOR Data[29]) XOR Data[48]) XOR Data[2]))) OR Data[11]);
    OutReady := 1;
    CollectInput(RESET:=TRUE);
  END_IF;
END_PROGRAM

CONFIGURATION Config0
  RESOURCE Res0 ON PLC
    TASK task0(INTERVAL := T#20ms,PRIORITY := 0);
    PROGRAM instance0 WITH task0 : Boiler;
  END_RESOURCE
END_CONFIGURATION

(* ---- RND-EXPR_bedew-mange-cater.st ---- *)
(*
This code implements a randomly grown symbolic expression:

xor(xor(((IN24 & (!(!(!(!((xor(xor(IN2, IN14), IN42)) & (!(IN8)))))))) | (!(!(!(IN31))))) | (xor(xor(((!((xor(xor((!(IN48)) | IN14, (xor(xor(IN19, IN16), IN34)) | IN30), (IN21 & IN10) & (IN24 | IN42))) & ((!(IN18)) | (xor(xor(IN48 | IN26, IN13 & IN15), xor(xor(IN39, IN12), IN50)))))) | ((!(xor(xor(!(xor(xor(IN49, IN23), IN44)), (!(IN11)) | (IN19 & IN50)), (!(IN17)) | IN32))) | ((xor(xor(IN22, IN12), xor(xor(!(IN35), !(IN5)), true))) | ((xor(xor(IN6 & IN2, IN32 | IN31), !(IN25))) | (!(IN39 & IN31)))))) | ((!(IN36)) | (!((!((IN35 | IN29) | (!(IN6)))) | IN42))), xor(xor(IN30, !(((xor(xor((IN5 & IN7) | IN29, (!(IN3)) | (IN47 & IN30)), IN2 & IN19)) | (((xor(xor(IN31, IN32), IN37)) | IN41) | (!(xor(xor(IN21, IN32), IN43))))) | IN15)), ((xor(xor(xor(xor(xor(xor(IN47, !(IN39)), IN19 & IN23), !(xor(xor(IN27, IN7), IN23))), (!(IN22)) & (!(IN40))), IN48 & ((IN50 | IN19) & (IN47 | IN3))), ((IN32 | IN4) | (IN17 & IN30)) & IN37)) | (!(!(IN50)))) & IN14)), IN41 & ((IN25 | ((((!(IN1)) & (IN14 | IN42)) | IN34) | ((!(xor(xor(IN8, IN37), IN49))) & (xor(xor(IN47, xor(xor(IN47, IN25), IN41)), !(IN37)))))) | ((((xor(xor(IN9, !(IN1)), IN6 & IN49)) | (xor(xor(xor(xor(IN11, false), IN4), IN31 | IN5), IN43 | IN9))) & (!(xor(xor(xor(xor(IN19, true), IN44), xor(xor(IN42, IN30), IN15)), IN18 | IN23)))) | ((xor(xor(!(IN5), (IN19 & IN29) | (IN13 & IN17)), (IN18 & IN44) & (xor(xor(IN31, IN31), IN16)))) | (IN22 | ((IN33 & IN41) | IN2))))))), (!(IN3)) & ((!(xor(xor((xor(xor((!(IN16 | IN16)) | (IN10 | (xor(xor(IN5, IN43), IN37))), !((xor(xor(IN20, IN7), IN23)) & (IN44 & IN19))), !((IN5 | IN25) | (IN31 & IN25)))) | (xor(xor((!(IN49 | IN12)) | ((!(IN37)) & (IN24 | false)), xor(xor(!(IN33 & IN45), !(IN49)), (xor(xor(IN12, IN27), IN49)) & (!(IN16)))), (xor(xor(IN43 & IN19, IN11 | IN50), IN29)) & IN34)), !(IN39)), xor(xor(!(IN35), true & ((!(!(IN2))) | ((xor(xor(IN35, IN32), IN44)) & (xor(xor(IN31, IN31), IN33))))), (!((xor(xor(IN1, IN12), IN49)) & (xor(xor(IN7, IN36), IN22)))) | (((IN49 & IN48) | (IN44 & IN4)) | (xor(xor(IN23 | IN1, xor(xor(IN24, IN20), IN10)), IN14 | IN45))))))) & ((!(IN42)) & IN31))), IN6)

*)

FUNCTION_BLOCK F_CollectInput
  VAR_IN_OUT
      Data : ARRAY[1..50] OF BOOL;
  END_VAR
  VAR_INPUT
      TICK  : BOOL := 0;
      IN1   : BOOL := 0;
      IN2   : BOOL := 0;
      IN3   : BOOL := 0;
      IN4   : BOOL := 0;
      IN5   : BOOL := 0;
      RESET : BOOL := FALSE;
  END_VAR
  VAR_OUTPUT
      Finished : BOOL;
  END_VAR
  VAR
      j    : USINT := 1;
      tock : BOOL  := 0;
  END_VAR
  IF NOT RESET AND tock = NOT TICK THEN
      Data[j]   := IN1;
      Data[j+1] := IN2;
      Data[j+2] := IN3;
      Data[j+3] := IN4;
      Data[j+4] := IN5;
      j := j + 5;
      tock := TICK;
  ELSE
      j := 1;
      tock := 0;
  END_IF;
  Finished := (j > 50);
END_FUNCTION_BLOCK

PROGRAM Boiler
  VAR
    Data  : ARRAY[1..50] OF BOOL;
    Ready : BOOL;
    CollectInput : F_CollectInput;
  END_VAR
  VAR
    TICK     AT %IX1.0 : BOOL;
    IN1      AT %IX0.3 : BOOL;
    IN2      AT %IX0.4 : BOOL;
    IN3      AT %IX0.5 : BOOL;
    IN4      AT %IX0.6 : BOOL;
    IN5      AT %IX0.7 : BOOL;
    OutReady AT %QX0.0 : BOOL := FALSE;
    FeedNext AT %QX0.1 : BOOL := FALSE;
    Out      AT %QX0.2 : BOOL;
  END_VAR
  CollectInput(TICK:=TICK, IN1:=IN1, IN2:=IN2, IN3:=IN3, IN4:=IN4, IN5:=IN5);
  Ready := CollectInput.Finished;
  FeedNext := 1;
  IF Ready THEN
    Out := (((((Data[24] AND (NOT (NOT (NOT (NOT (((Data[2] XOR Data[14]) XOR Data[42]) AND (NOT Data[8]))))))) OR (NOT (NOT (NOT Data[31])))) OR (((((NOT (((((NOT Data[48]) OR Data[14]) XOR (((Data[19] XOR Data[16]) XOR Data[34]) OR Data[30])) XOR ((Data[21] AND Data[10]) AND (Data[24] OR Data[42]))) AND ((NOT Data[18]) OR (((Data[48] OR Data[26]) XOR (Data[13] AND Data[15])) XOR ((Data[39] XOR Data[12]) XOR Data[50]))))) OR ((NOT (((NOT ((Data[49] XOR Data[23]) XOR Data[44])) XOR ((NOT Data[11]) OR (Data[19] AND Data[50]))) XOR ((NOT Data[17]) OR Data[32]))) OR (((Data[22] XOR Data[12]) XOR (((NOT Data[35]) XOR (NOT Data[5])) XOR TRUE)) OR ((((Data[6] AND Data[2]) XOR (Data[32] OR Data[31])) XOR (NOT Data[25])) OR (NOT (Data[39] AND Data[31])))))) OR ((NOT Data[36]) OR (NOT ((NOT ((Data[35] OR Data[29]) OR (NOT Data[6]))) OR Data[42])))) XOR ((Data[30] XOR (NOT ((((((Data[5] AND Data[7]) OR Data[29]) XOR ((NOT Data[3]) OR (Data[47] AND Data[30]))) XOR (Data[2] AND Data[19])) OR ((((Data[31] XOR Data[32]) XOR Data[37]) OR Data[41]) OR (NOT ((Data[21] XOR Data[32]) XOR Data[43])))) OR Data[15]))) XOR ((((((((Data[47] XOR (NOT Data[39])) XOR (Data[19] AND Data[23])) XOR (NOT ((Data[27] XOR Data[7]) XOR Data[23]))) XOR ((NOT Data[22]) AND (NOT Data[40]))) XOR (Data[48] AND ((Data[50] OR Data[19]) AND (Data[47] OR Data[3])))) XOR (((Data[32] OR Data[4]) OR (Data[17] AND Data[30])) AND Data[37])) OR (NOT (NOT Data[50]))) AND Data[14]))) XOR (Data[41] AND ((Data[25] OR ((((NOT Data[1]) AND (Data[14] OR Data[42])) OR Data[34]) OR ((NOT ((Data[8] XOR Data[37]) XOR Data[49])) AND ((Data[47] XOR ((Data[47] XOR Data[25]) XOR Data[41])) XOR (NOT Data[37]))))) OR (((((Data[9] XOR (NOT Data[1])) XOR (Data[6] AND Data[49])) OR ((((Data[11] XOR FALSE) XOR Data[4]) XOR (Data[31] OR Data[5])) XOR (Data[43] OR Data[9]))) AND (NOT ((((Data[19] XOR TRUE) XOR Data[44]) XOR ((Data[42] XOR Data[30]) XOR Data[15])) XOR (Data[18] OR Data[23])))) OR ((((NOT Data[5]) XOR ((Data[19] AND Data[29]) OR (Data[13] AND Data[17]))) XOR ((Data[18] AND Data[44]) AND ((Data[31] XOR Data[31]) XOR Data[16]))) OR (Data[22] OR ((Data[33] AND Data[41]) OR Data[2])))))))) XOR ((NOT Data[3]) AND ((NOT (((((((NOT (Data[16] OR Data[16])) OR (Data[10] OR ((Data[5] XOR Data[43]) XOR Data[37]))) XOR (NOT (((Data[20] XOR Data[7]) XOR Data[23]) AND (Data[44] AND Data[19])))) XOR (NOT ((Data[5] OR Data[25]) OR (Data[31] AND Data[25])))) OR ((((NOT (Data[49] OR Data[12])) OR ((NOT Data[37]) AND (Data[24] OR FALSE))) XOR (((NOT (Data[33] AND Data[45])) XOR (NOT Data[49])) XOR (((Data[12] XOR Data[27]) XOR Data[49]) AND (NOT Data[16])))) XOR ((((Data[43] AND Data[19]) XOR (Data[11] OR Data[50])) XOR Data[29]) AND Data[34]))) XOR (NOT Data[39])) XOR (((NOT Data[35]) XOR (TRUE AND ((NOT (NOT Data[2])) OR (((Data[35] XOR Data[32]) XOR Data[44]) AND ((Data[31] XOR Data[31]) XOR Data[33]))))) XOR ((NOT (((Data[1] XOR Data[12]) XOR Data[49]) AND ((Data[7] XOR Data[36]) XOR Data[22]))) OR (((Data[49] AND Data[48]) OR (Data[44] AND Data[4])) OR (((Data[23] OR Data[1]) XOR ((Data[24] XOR Data[20]) XOR Data[10])) XOR (Data[14] OR Data[45]))))))) AND ((NOT Data[42]) AND Data[31])))) XOR Data[6]);
    OutReady := 1;
    CollectInput(RESET:=TRUE);
  END_IF;
END_PROGRAM

CONFIGURATION Config0
  RESOURCE Res0 ON PLC
    TASK task0(INTERVAL := T#20ms,PRIORITY := 0);
    PROGRAM instance0 WITH task0 : Boiler;
  END_RESOURCE
END_CONFIGURATION

(* ---- RND-EXPR_belay-palsy-rifts.st ---- *)
(*
This code implements a randomly grown symbolic expression:

xor(xor((IN16 | IN26) & ((((xor(xor(!(xor(xor(IN38 | (!(IN38)), !(!(IN8))), !(xor(xor(IN44, IN37), IN27)))), (((!(IN1)) & (IN27 | IN45)) | (IN40 & (IN38 & IN27))) & IN36), ((!(!(IN43))) | ((xor(xor(IN16, IN18), IN25)) & (IN45 & IN43))) & (((!(IN16)) | (IN31 & IN9)) & (xor(xor(IN8, IN40), IN38 | IN17))))) & (xor(xor(((!(IN27)) & ((!(IN1)) | (IN35 & IN28))) | ((!(!(IN15))) & IN32), (((IN48 & IN5) | (IN10 | true)) | true) | (xor(xor(false, !(xor(xor(IN43, IN3), IN44))), xor(xor(xor(xor(IN49, IN34), IN16), IN12 | IN26), IN6)))), (IN39 & (xor(xor(IN46 & IN10, IN22 | IN11), xor(xor(IN46, IN12), true)))) | IN28))) | (!((xor(xor(xor(xor((IN45 | IN44) | (IN15 | IN13), (!(IN36)) | (IN45 | IN39)), !(IN9 & IN49)), (xor(xor(xor(xor(IN4, IN37), IN21), xor(xor(IN9, IN19), IN3)), IN30 & IN16)) | (!(xor(xor(IN25, IN45), IN33)))), ((IN40 & IN16) | (!(IN39))) | ((xor(xor(IN25, IN35), IN21)) & (IN30 & IN29)))) | (xor(xor(IN16, (!(IN5 & IN15)) | (!(!(IN18)))), IN49))))) & (IN39 | (!(((IN38 & IN11) & (!((!(IN25)) | (!(IN2))))) | IN25)))), IN25), IN6 & ((!(xor(xor(!(xor(xor(xor(xor((xor(xor(IN45, IN32), IN43)) & (IN9 | IN44), false), xor(xor(IN13 | IN25, IN9 & IN14), IN48 | IN42)), !((!(IN11)) & (!(IN27)))), (!(IN25)) | (!(!(IN48))))), (!(IN15)) | (xor(xor(xor(xor((xor(xor(IN48, false), IN4)) & (xor(xor(IN34, IN46), IN33)), !(xor(xor(IN7, IN46), IN31))), xor(xor(!(IN13), false & IN43), xor(xor(IN13, IN36), IN26))), ((false | IN10) | (IN24 | IN15)) & IN38), IN14 | (xor(xor(IN50, xor(xor(IN3, IN1), IN14)), !(IN43)))))), !((xor(xor(!(xor(xor(IN23, false), IN25)), xor(xor(xor(xor(IN21, IN7), IN18), IN32 | IN34), xor(xor(IN28, IN2), IN43))), IN35)) | (((!(IN47)) & (IN50 | IN28)) | (xor(xor(IN45 | IN1, IN16 & IN45), IN29))))))) & (xor(xor(!(xor(xor(xor(xor(IN32, xor(xor(!(IN42 & IN4), IN22), IN42 & (!(IN46)))), xor(xor(IN6, (!(IN37)) | (IN11 & IN40)), (!(IN50)) | (false & IN45))), !((IN20 | (!(IN44))) & IN32)), !(((xor(xor(IN19, IN36), IN22)) | (IN38 & IN45)) & (!(!(IN35)))))), xor(xor(!(IN34), (!(IN3)) | IN50), !((xor(xor((IN16 | IN18) & IN41, xor(xor(IN50, xor(xor(IN2, IN44), IN23)), xor(xor(IN8, IN43), IN19))), xor(xor(IN11 | IN29, !(IN44)), !(IN27)))) | IN45))), (!((!(IN30 | (xor(xor(IN45, IN14), IN20)))) & (xor(xor(!(IN18), (IN13 | false) & (IN8 & IN46)), IN28)))) | IN20))))

*)

FUNCTION_BLOCK F_CollectInput
  VAR_IN_OUT
      Data : ARRAY[1..50] OF BOOL;
  END_VAR
  VAR_INPUT
      TICK  : BOOL := 0;
      IN1   : BOOL := 0;
      IN2   : BOOL := 0;
      IN3   : BOOL := 0;
      IN4   : BOOL := 0;
      IN5   : BOOL := 0;
      RESET : BOOL := FALSE;
  END_VAR
  VAR_OUTPUT
      Finished : BOOL;
  END_VAR
  VAR
      j    : USINT := 1;
      tock : BOOL  := 0;
  END_VAR
  IF NOT RESET AND tock = NOT TICK THEN
      Data[j]   := IN1;
      Data[j+1] := IN2;
      Data[j+2] := IN3;
      Data[j+3] := IN4;
      Data[j+4] := IN5;
      j := j + 5;
      tock := TICK;
  ELSE
      j := 1;
      tock := 0;
  END_IF;
  Finished := (j > 50);
END_FUNCTION_BLOCK

PROGRAM Boiler
  VAR
    Data  : ARRAY[1..50] OF BOOL;
    Ready : BOOL;
    CollectInput : F_CollectInput;
  END_VAR
  VAR
    TICK     AT %IX1.0 : BOOL;
    IN1      AT %IX0.3 : BOOL;
    IN2      AT %IX0.4 : BOOL;
    IN3      AT %IX0.5 : BOOL;
    IN4      AT %IX0.6 : BOOL;
    IN5      AT %IX0.7 : BOOL;
    OutReady AT %QX0.0 : BOOL := FALSE;
    FeedNext AT %QX0.1 : BOOL := FALSE;
    Out      AT %QX0.2 : BOOL;
  END_VAR
  CollectInput(TICK:=TICK, IN1:=IN1, IN2:=IN2, IN3:=IN3, IN4:=IN4, IN5:=IN5);
  Ready := CollectInput.Finished;
  FeedNext := 1;
  IF Ready THEN
    Out := ((((Data[16] OR Data[26]) AND ((((((NOT (((Data[38] OR (NOT Data[38])) XOR (NOT (NOT Data[8]))) XOR (NOT ((Data[44] XOR Data[37]) XOR Data[27])))) XOR ((((NOT Data[1]) AND (Data[27] OR Data[45])) OR (Data[40] AND (Data[38] AND Data[27]))) AND Data[36])) XOR (((NOT (NOT Data[43])) OR (((Data[16] XOR Data[18]) XOR Data[25]) AND (Data[45] AND Data[43]))) AND (((NOT Data[16]) OR (Data[31] AND Data[9])) AND ((Data[8] XOR Data[40]) XOR (Data[38] OR Data[17]))))) AND (((((NOT Data[27]) AND ((NOT Data[1]) OR (Data[35] AND Data[28]))) OR ((NOT (NOT Data[15])) AND Data[32])) XOR ((((Data[48] AND Data[5]) OR (Data[10] OR TRUE)) OR TRUE) OR ((FALSE XOR (NOT ((Data[43] XOR Data[3]) XOR Data[44]))) XOR ((((Data[49] XOR Data[34]) XOR Data[16]) XOR (Data[12] OR Data[26])) XOR Data[6])))) XOR ((Data[39] AND (((Data[46] AND Data[10]) XOR (Data[22] OR Data[11])) XOR ((Data[46] XOR Data[12]) XOR TRUE))) OR Data[28]))) OR (NOT (((((((Data[45] OR Data[44]) OR (Data[15] OR Data[13])) XOR ((NOT Data[36]) OR (Data[45] OR Data[39]))) XOR (NOT (Data[9] AND Data[49]))) XOR (((((Data[4] XOR Data[37]) XOR Data[21]) XOR ((Data[9] XOR Data[19]) XOR Data[3])) XOR (Data[30] AND Data[16])) OR (NOT ((Data[25] XOR Data[45]) XOR Data[33])))) XOR (((Data[40] AND Data[16]) OR (NOT Data[39])) OR (((Data[25] XOR Data[35]) XOR Data[21]) AND (Data[30] AND Data[29])))) OR ((Data[16] XOR ((NOT (Data[5] AND Data[15])) OR (NOT (NOT Data[18])))) XOR Data[49])))) AND (Data[39] OR (NOT (((Data[38] AND Data[11]) AND (NOT ((NOT Data[25]) OR (NOT Data[2])))) OR Data[25]))))) XOR Data[25]) XOR (Data[6] AND ((NOT (((NOT (((((((Data[45] XOR Data[32]) XOR Data[43]) AND (Data[9] OR Data[44])) XOR FALSE) XOR (((Data[13] OR Data[25]) XOR (Data[9] AND Data[14])) XOR (Data[48] OR Data[42]))) XOR (NOT ((NOT Data[11]) AND (NOT Data[27])))) XOR ((NOT Data[25]) OR (NOT (NOT Data[48]))))) XOR ((NOT Data[15]) OR (((((((Data[48] XOR FALSE) XOR Data[4]) AND ((Data[34] XOR Data[46]) XOR Data[33])) XOR (NOT ((Data[7] XOR Data[46]) XOR Data[31]))) XOR (((NOT Data[13]) XOR (FALSE AND Data[43])) XOR ((Data[13] XOR Data[36]) XOR Data[26]))) XOR (((FALSE OR Data[10]) OR (Data[24] OR Data[15])) AND Data[38])) XOR (Data[14] OR ((Data[50] XOR ((Data[3] XOR Data[1]) XOR Data[14])) XOR (NOT Data[43])))))) XOR (NOT ((((NOT ((Data[23] XOR FALSE) XOR Data[25])) XOR ((((Data[21] XOR Data[7]) XOR Data[18]) XOR (Data[32] OR Data[34])) XOR ((Data[28] XOR Data[2]) XOR Data[43]))) XOR Data[35]) OR (((NOT Data[47]) AND (Data[50] OR Data[28])) OR (((Data[45] OR Data[1]) XOR (Data[16] AND Data[45])) XOR Data[29])))))) AND (((NOT ((((Data[32] XOR (((NOT (Data[42] AND Data[4])) XOR Data[22]) XOR (Data[42] AND (NOT Data[46])))) XOR ((Data[6] XOR ((NOT Data[37]) OR (Data[11] AND Data[40]))) XOR ((NOT Data[50]) OR (FALSE AND Data[45])))) XOR (NOT ((Data[20] OR (NOT Data[44])) AND Data[32]))) XOR (NOT ((((Data[19] XOR Data[36]) XOR Data[22]) OR (Data[38] AND Data[45])) AND (NOT (NOT Data[35])))))) XOR (((NOT Data[34]) XOR ((NOT Data[3]) OR Data[50])) XOR (NOT (((((Data[16] OR Data[18]) AND Data[41]) XOR ((Data[50] XOR ((Data[2] XOR Data[44]) XOR Data[23])) XOR ((Data[8] XOR Data[43]) XOR Data[19]))) XOR (((Data[11] OR Data[29]) XOR (NOT Data[44])) XOR (NOT Data[27]))) OR Data[45])))) XOR ((NOT ((NOT (Data[30] OR ((Data[45] XOR Data[14]) XOR Data[20]))) AND (((NOT Data[18]) XOR ((Data[13] OR FALSE) AND (Data[8] AND Data[46]))) XOR Data[28]))) OR Data[20])))));
    OutReady := 1;
    CollectInput(RESET:=TRUE);
  END_IF;
END_PROGRAM

CONFIGURATION Config0
  RESOURCE Res0 ON PLC
    TASK task0(INTERVAL := T#20ms,PRIORITY := 0);
    PROGRAM instance0 WITH task0 : Boiler;
  END_RESOURCE
END_CONFIGURATION

(* ---- RND-EXPR_birch-anole-elope.st ---- *)
(*
This code implements a randomly grown symbolic expression:

(xor(xor(!(!(xor(xor(xor(xor((IN6 | ((IN4 & IN40) | true)) | IN7, xor(xor(!(IN4), IN38 & IN9), xor(xor(!(!(IN39)), !(IN9)), (IN20 & IN48) & IN8))), xor(xor(IN49, IN49), xor(xor((xor(xor(IN3, true), IN17)) & (xor(xor(IN50, IN27), IN18)), IN17 | IN24), (xor(xor(IN5, IN32), IN45)) & (xor(xor(IN23, IN35), IN16))))), (IN48 & (IN1 | ((true | IN6) | IN50))) & IN23), true))), !(!(IN36 | (IN23 | (!(!(xor(xor(!(IN21), IN9 & IN45), IN50 & IN23)))))))), xor(xor(!((!(!(xor(xor(!(xor(xor(IN14, IN48), IN22)), !(IN31 | IN8)), IN42 | (false | IN43))))) & IN24), !(xor(xor(xor(xor(IN6 & (((!(IN33)) | (!(IN34))) | ((IN28 | false) | IN6)), IN4), ((xor(xor(true, IN2 & IN24), !(IN40))) & (IN33 & (xor(xor(IN16, IN17), IN30)))) & ((!(IN9)) | IN10)), IN19 & (xor(xor(IN43, (xor(xor(!(IN20), IN23 & IN40), IN4 | IN34)) | ((!(IN3)) & (IN28 | IN13))), ((IN38 & IN26) & (IN23 & IN41)) | ((IN47 | IN39) & (xor(xor(IN28, IN31), IN9)))))), IN24 | (xor(xor(((IN44 | IN34) & (!(IN15))) | (IN8 | IN30), !(IN24)), !(xor(xor(IN1 | IN15, IN37 & IN22), IN34))))))), (!(!(IN3))) | ((!((!(!(IN41 & IN5))) | (((IN15 & IN30) | (!(IN41))) & (!(xor(xor(IN45, IN23), IN49)))))) | (!((IN15 & (xor(xor(IN33, IN35 | IN31), IN17 | IN11))) & ((!(IN48)) & ((!(IN43)) & (IN5 | IN43))))))))) | ((xor(xor(xor(xor(!(IN1), IN16 | IN9), !(IN31)), IN3), (((xor(xor(!(xor(xor(xor(xor(IN26, IN1), IN8), IN16 | IN23), IN27)), xor(xor(IN48 & (xor(xor(IN25, IN21), IN45)), IN24), !(IN37 & IN25))), ((IN34 & IN27) | IN11) | (xor(xor(IN48, xor(xor(IN50, IN12), IN35)), !(IN24))))) & (IN20 | (((xor(xor(IN43, IN17), IN24)) | (!(IN15))) & IN18))) & (IN17 & (!(IN41)))) | (!(xor(xor((IN39 | (xor(xor(!(IN19), IN39 & IN47), xor(xor(IN18, IN45), IN1)))) | (xor(xor((false & IN8) & (IN7 & IN19), !(IN39 & IN17)), !(!(IN44)))), (((IN4 | IN27) | IN8) & (!(!(IN38)))) | (IN48 | (xor(xor(!(IN18), xor(xor(IN18, IN41), IN36)), IN42 | IN14)))), IN21))))) & ((!(!(IN1))) & (!((xor(xor(xor(xor(xor(xor((IN38 | IN1) | (IN13 & IN33), (!(IN17)) & (IN12 & IN16)), (!(IN39)) | (!(IN41))), (!(IN43 | IN4)) & (xor(xor(xor(xor(IN2, IN6), IN8), xor(xor(IN33, IN43), IN22)), true & IN25))), IN41 | ((IN43 | IN46) & (IN10 & IN14))), (!(!(IN42 & IN34))) | IN29), !(((!(IN49)) & (IN33 & IN20)) | (xor(xor(IN1, IN19 | IN21), IN12))))) | ((xor(xor(!((!(IN32)) & (!(IN44))), IN21 & (xor(xor(IN35 | IN42, xor(xor(IN34, IN17), IN1)), IN49 & IN37))), ((!(IN15)) & IN30) & (xor(xor(false, IN37 & IN31), IN42)))) & ((((!(IN36)) & IN22) & (xor(xor(IN48, IN37 & IN48), IN13))) | (xor(xor(IN8 & IN42, IN40), false))))))))

*)

FUNCTION_BLOCK F_CollectInput
  VAR_IN_OUT
      Data : ARRAY[1..50] OF BOOL;
  END_VAR
  VAR_INPUT
      TICK  : BOOL := 0;
      IN1   : BOOL := 0;
      IN2   : BOOL := 0;
      IN3   : BOOL := 0;
      IN4   : BOOL := 0;
      IN5   : BOOL := 0;
      RESET : BOOL := FALSE;
  END_VAR
  VAR_OUTPUT
      Finished : BOOL;
  END_VAR
  VAR
      j    : USINT := 1;
      tock : BOOL  := 0;
  END_VAR
  IF NOT RESET AND tock = NOT TICK THEN
      Data[j]   := IN1;
      Data[j+1] := IN2;
      Data[j+2] := IN3;
      Data[j+3] := IN4;
      Data[j+4] := IN5;
      j := j + 5;
      tock := TICK;
  ELSE
      j := 1;
      tock := 0;
  END_IF;
  Finished := (j > 50);
END_FUNCTION_BLOCK

PROGRAM Boiler
  VAR
    Data  : ARRAY[1..50] OF BOOL;
    Ready : BOOL;
    CollectInput : F_CollectInput;
  END_VAR
  VAR
    TICK     AT %IX1.0 : BOOL;
    IN1      AT %IX0.3 : BOOL;
    IN2      AT %IX0.4 : BOOL;
    IN3      AT %IX0.5 : BOOL;
    IN4      AT %IX0.6 : BOOL;
    IN5      AT %IX0.7 : BOOL;
    OutReady AT %QX0.0 : BOOL := FALSE;
    FeedNext AT %QX0.1 : BOOL := FALSE;
    Out      AT %QX0.2 : BOOL;
  END_VAR
  CollectInput(TICK:=TICK, IN1:=IN1, IN2:=IN2, IN3:=IN3, IN4:=IN4, IN5:=IN5);
  Ready := CollectInput.Finished;
  FeedNext := 1;
  IF Ready THEN
    Out := ((((NOT (NOT ((((((Data[6] OR ((Data[4] AND Data[40]) OR TRUE)) OR Data[7]) XOR (((NOT Data[4]) XOR (Data[38] AND Data[9])) XOR (((NOT (NOT Data[39])) XOR (NOT Data[9])) XOR ((Data[20] AND Data[48]) AND Data[8])))) XOR ((Data[49] XOR Data[49]) XOR (((((Data[3] XOR TRUE) XOR Data[17]) AND ((Data[50] XOR Data[27]) XOR Data[18])) XOR (Data[17] OR Data[24])) XOR (((Data[5] XOR Data[32]) XOR Data[45]) AND ((Data[23] XOR Data[35]) XOR Data[16]))))) XOR ((Data[48] AND (Data[1] OR ((TRUE OR Data[6]) OR Data[50]))) AND Data[23])) XOR TRUE))) XOR (NOT (NOT (Data[36] OR (Data[23] OR (NOT (NOT (((NOT Data[21]) XOR (Data[9] AND Data[45])) XOR (Data[50] AND Data[23]))))))))) XOR (((NOT ((NOT (NOT (((NOT ((Data[14] XOR Data[48]) XOR Data[22])) XOR (NOT (Data[31] OR Data[8]))) XOR (Data[42] OR (FALSE OR Data[43]))))) AND Data[24])) XOR (NOT (((((Data[6] AND (((NOT Data[33]) OR (NOT Data[34])) OR ((Data[28] OR FALSE) OR Data[6]))) XOR Data[4]) XOR ((((TRUE XOR (Data[2] AND Data[24])) XOR (NOT Data[40])) AND (Data[33] AND ((Data[16] XOR Data[17]) XOR Data[30]))) AND ((NOT Data[9]) OR Data[10]))) XOR (Data[19] AND ((Data[43] XOR ((((NOT Data[20]) XOR (Data[23] AND Data[40])) XOR (Data[4] OR Data[34])) OR ((NOT Data[3]) AND (Data[28] OR Data[13])))) XOR (((Data[38] AND Data[26]) AND (Data[23] AND Data[41])) OR ((Data[47] OR Data[39]) AND ((Data[28] XOR Data[31]) XOR Data[9])))))) XOR (Data[24] OR (((((Data[44] OR Data[34]) AND (NOT Data[15])) OR (Data[8] OR Data[30])) XOR (NOT Data[24])) XOR (NOT (((Data[1] OR Data[15]) XOR (Data[37] AND Data[22])) XOR Data[34]))))))) XOR ((NOT (NOT Data[3])) OR ((NOT ((NOT (NOT (Data[41] AND Data[5]))) OR (((Data[15] AND Data[30]) OR (NOT Data[41])) AND (NOT ((Data[45] XOR Data[23]) XOR Data[49]))))) OR (NOT ((Data[15] AND ((Data[33] XOR (Data[35] OR Data[31])) XOR (Data[17] OR Data[11]))) AND ((NOT Data[48]) AND ((NOT Data[43]) AND (Data[5] OR Data[43]))))))))) OR ((((((NOT Data[1]) XOR (Data[16] OR Data[9])) XOR (NOT Data[31])) XOR Data[3]) XOR ((((((NOT ((((Data[26] XOR Data[1]) XOR Data[8]) XOR (Data[16] OR Data[23])) XOR Data[27])) XOR (((Data[48] AND ((Data[25] XOR Data[21]) XOR Data[45])) XOR Data[24]) XOR (NOT (Data[37] AND Data[25])))) XOR (((Data[34] AND Data[27]) OR Data[11]) OR ((Data[48] XOR ((Data[50] XOR Data[12]) XOR Data[35])) XOR (NOT Data[24])))) AND (Data[20] OR ((((Data[43] XOR Data[17]) XOR Data[24]) OR (NOT Data[15])) AND Data[18]))) AND (Data[17] AND (NOT Data[41]))) OR (NOT ((((Data[39] OR (((NOT Data[19]) XOR (Data[39] AND Data[47])) XOR ((Data[18] XOR Data[45]) XOR Data[1]))) OR ((((FALSE AND Data[8]) AND (Data[7] AND Data[19])) XOR (NOT (Data[39] AND Data[17]))) XOR (NOT (NOT Data[44])))) XOR ((((Data[4] OR Data[27]) OR Data[8]) AND (NOT (NOT Data[38]))) OR (Data[48] OR (((NOT Data[18]) XOR ((Data[18] XOR Data[41]) XOR Data[36])) XOR (Data[42] OR Data[14]))))) XOR Data[21])))) AND ((NOT (NOT Data[1])) AND (NOT (((((((((Data[38] OR Data[1]) OR (Data[13] AND Data[33])) XOR ((NOT Data[17]) AND (Data[12] AND Data[16]))) XOR ((NOT Data[39]) OR (NOT Data[41]))) XOR ((NOT (Data[43] OR Data[4])) AND ((((Data[2] XOR Data[6]) XOR Data[8]) XOR ((Data[33] XOR Data[43]) XOR Data[22])) XOR (TRUE AND Data[25])))) XOR (Data[41] OR ((Data[43] OR Data[46]) AND (Data[10] AND Data[14])))) XOR ((NOT (NOT (Data[42] AND Data[34]))) OR Data[29])) XOR (NOT (((NOT Data[49]) AND (Data[33] AND Data[20])) OR ((Data[1] XOR (Data[19] OR Data[21])) XOR Data[12])))) OR ((((NOT ((NOT Data[32]) AND (NOT Data[44]))) XOR (Data[21] AND (((Data[35] OR Data[42]) XOR ((Data[34] XOR Data[17]) XOR Data[1])) XOR (Data[49] AND Data[37])))) XOR (((NOT Data[15]) AND Data[30]) AND ((FALSE XOR (Data[37] AND Data[31])) XOR Data[42]))) AND ((((NOT Data[36]) AND Data[22]) AND ((Data[48] XOR (Data[37] AND Data[48])) XOR Data[13])) OR (((Data[8] AND Data[42]) XOR Data[40]) XOR FALSE))))))));
    OutReady := 1;
    CollectInput(RESET:=TRUE);
  END_IF;
END_PROGRAM

CONFIGURATION Config0
  RESOURCE Res0 ON PLC
    TASK task0(INTERVAL := T#20ms,PRIORITY := 0);
    PROGRAM instance0 WITH task0 : Boiler;
  END_RESOURCE
END_CONFIGURATION

(* ---- RND-EXPR_bland-kicky-recto.st ---- *)
(*
This code implements a randomly grown symbolic expression:

((xor(xor(xor(xor(xor(xor(IN48, xor(xor((!((xor(xor(IN5, IN42), IN45)) | (IN37 & false))) & (xor(xor(xor(xor(IN2, !(IN14)), IN48), xor(xor(IN21 | IN17, IN27 | IN19), IN36)), !(IN13 & IN45))), IN27), ((!(xor(xor(IN17, IN29), IN43))) & ((xor(xor(IN39, IN3), IN34)) | IN14)) & ((!(xor(xor(IN39, IN41), IN17))) & true))), IN46), !(!((IN43 & ((xor(xor(IN37, IN8), IN48)) & (IN16 & IN16))) & (!((IN15 | IN18) | IN37))))), (xor(xor(!(IN34 & (xor(xor(IN9 & IN18, xor(xor(false, IN44), IN30)), IN5))), xor(xor(((!(IN48)) | (IN17 & IN37)) | IN1, !((xor(xor(IN10, IN18), IN41)) | (IN45 & IN13))), IN4 | (!(IN41 & IN27)))), !((!(IN7 | IN36)) & ((!(IN20)) | IN9)))) | ((!(!(IN29))) | IN6)), IN2), xor(xor(IN43 | (xor(xor(((xor(xor(!(IN14), !(IN15)), xor(xor(IN1, IN15), IN50))) & ((IN10 & IN6) & (IN6 | IN7))) | (!((IN15 | IN26) | (!(IN41)))), xor(xor(!(!(!(IN43))), IN36 & IN15), IN31 | (IN42 & (IN48 & IN47)))), ((xor(xor(!(IN23), IN15 & IN10), IN31)) & (xor(xor(xor(xor(IN29, IN46), false), IN15), !(IN7)))) & IN24)), xor(xor(IN5, IN16), !((!(!(xor(xor(IN10, IN47), IN10)))) | (IN8 | ((!(IN18)) | (!(IN31))))))), (true | ((!(xor(xor(IN20 | IN43, IN4 & IN11), !(IN3)))) | (IN17 | (!(IN28 | IN3))))) | ((!(!((IN18 | IN37) & (xor(xor(IN12, IN43), IN4))))) & IN23)))) & ((!(IN17)) & (!(IN45)))) | (IN33 & (xor(xor(!(IN17), xor(xor(!((xor(xor(!(!(!(IN39))), xor(xor(!(IN13 & IN33), IN33 | IN16), (xor(xor(IN3, IN11), IN19)) & (IN6 | IN22))), ((IN18 & IN3) | (IN40 | IN23)) | ((IN41 | true) & IN44))) & IN13), (!(IN9 & (((!(IN38)) | (true & IN36)) & IN38))) & (!(((!(!(IN46))) & ((IN15 & IN28) & (IN16 | IN9))) & ((xor(xor(IN7, !(IN13)), IN41 & IN6)) | (xor(xor(xor(xor(IN40, IN31), IN6), !(IN39)), !(IN46))))))), IN11)), IN35)))

*)

FUNCTION_BLOCK F_CollectInput
  VAR_IN_OUT
      Data : ARRAY[1..50] OF BOOL;
  END_VAR
  VAR_INPUT
      TICK  : BOOL := 0;
      IN1   : BOOL := 0;
      IN2   : BOOL := 0;
      IN3   : BOOL := 0;
      IN4   : BOOL := 0;
      IN5   : BOOL := 0;
      RESET : BOOL := FALSE;
  END_VAR
  VAR_OUTPUT
      Finished : BOOL;
  END_VAR
  VAR
      j    : USINT := 1;
      tock : BOOL  := 0;
  END_VAR
  IF NOT RESET AND tock = NOT TICK THEN
      Data[j]   := IN1;
      Data[j+1] := IN2;
      Data[j+2] := IN3;
      Data[j+3] := IN4;
      Data[j+4] := IN5;
      j := j + 5;
      tock := TICK;
  ELSE
      j := 1;
      tock := 0;
  END_IF;
  Finished := (j > 50);
END_FUNCTION_BLOCK

PROGRAM Boiler
  VAR
    Data  : ARRAY[1..50] OF BOOL;
    Ready : BOOL;
    CollectInput : F_CollectInput;
  END_VAR
  VAR
    TICK     AT %IX1.0 : BOOL;
    IN1      AT %IX0.3 : BOOL;
    IN2      AT %IX0.4 : BOOL;
    IN3      AT %IX0.5 : BOOL;
    IN4      AT %IX0.6 : BOOL;
    IN5      AT %IX0.7 : BOOL;
    OutReady AT %QX0.0 : BOOL := FALSE;
    FeedNext AT %QX0.1 : BOOL := FALSE;
    Out      AT %QX0.2 : BOOL;
  END_VAR
  CollectInput(TICK:=TICK, IN1:=IN1, IN2:=IN2, IN3:=IN3, IN4:=IN4, IN5:=IN5);
  Ready := CollectInput.Finished;
  FeedNext := 1;
  IF Ready THEN
    Out := ((((((((Data[48] XOR ((((NOT (((Data[5] XOR Data[42]) XOR Data[45]) OR (Data[37] AND FALSE))) AND ((((Data[2] XOR (NOT Data[14])) XOR Data[48]) XOR (((Data[21] OR Data[17]) XOR (Data[27] OR Data[19])) XOR Data[36])) XOR (NOT (Data[13] AND Data[45])))) XOR Data[27]) XOR (((NOT ((Data[17] XOR Data[29]) XOR Data[43])) AND (((Data[39] XOR Data[3]) XOR Data[34]) OR Data[14])) AND ((NOT ((Data[39] XOR Data[41]) XOR Data[17])) AND TRUE)))) XOR Data[46]) XOR (NOT (NOT ((Data[43] AND (((Data[37] XOR Data[8]) XOR Data[48]) AND (Data[16] AND Data[16]))) AND (NOT ((Data[15] OR Data[18]) OR Data[37])))))) XOR ((((NOT (Data[34] AND (((Data[9] AND Data[18]) XOR ((FALSE XOR Data[44]) XOR Data[30])) XOR Data[5]))) XOR (((((NOT Data[48]) OR (Data[17] AND Data[37])) OR Data[1]) XOR (NOT (((Data[10] XOR Data[18]) XOR Data[41]) OR (Data[45] AND Data[13])))) XOR (Data[4] OR (NOT (Data[41] AND Data[27]))))) XOR (NOT ((NOT (Data[7] OR Data[36])) AND ((NOT Data[20]) OR Data[9])))) OR ((NOT (NOT Data[29])) OR Data[6]))) XOR Data[2]) XOR (((Data[43] OR (((((((NOT Data[14]) XOR (NOT Data[15])) XOR ((Data[1] XOR Data[15]) XOR Data[50])) AND ((Data[10] AND Data[6]) AND (Data[6] OR Data[7]))) OR (NOT ((Data[15] OR Data[26]) OR (NOT Data[41])))) XOR (((NOT (NOT (NOT Data[43]))) XOR (Data[36] AND Data[15])) XOR (Data[31] OR (Data[42] AND (Data[48] AND Data[47]))))) XOR (((((NOT Data[23]) XOR (Data[15] AND Data[10])) XOR Data[31]) AND ((((Data[29] XOR Data[46]) XOR FALSE) XOR Data[15]) XOR (NOT Data[7]))) AND Data[24]))) XOR ((Data[5] XOR Data[16]) XOR (NOT ((NOT (NOT ((Data[10] XOR Data[47]) XOR Data[10]))) OR (Data[8] OR ((NOT Data[18]) OR (NOT Data[31]))))))) XOR ((TRUE OR ((NOT (((Data[20] OR Data[43]) XOR (Data[4] AND Data[11])) XOR (NOT Data[3]))) OR (Data[17] OR (NOT (Data[28] OR Data[3]))))) OR ((NOT (NOT ((Data[18] OR Data[37]) AND ((Data[12] XOR Data[43]) XOR Data[4])))) AND Data[23])))) AND ((NOT Data[17]) AND (NOT Data[45]))) OR (Data[33] AND (((NOT Data[17]) XOR (((NOT ((((NOT (NOT (NOT Data[39]))) XOR (((NOT (Data[13] AND Data[33])) XOR (Data[33] OR Data[16])) XOR (((Data[3] XOR Data[11]) XOR Data[19]) AND (Data[6] OR Data[22])))) XOR (((Data[18] AND Data[3]) OR (Data[40] OR Data[23])) OR ((Data[41] OR TRUE) AND Data[44]))) AND Data[13])) XOR ((NOT (Data[9] AND (((NOT Data[38]) OR (TRUE AND Data[36])) AND Data[38]))) AND (NOT (((NOT (NOT Data[46])) AND ((Data[15] AND Data[28]) AND (Data[16] OR Data[9]))) AND (((Data[7] XOR (NOT Data[13])) XOR (Data[41] AND Data[6])) OR ((((Data[40] XOR Data[31]) XOR Data[6]) XOR (NOT Data[39])) XOR (NOT Data[46]))))))) XOR Data[11])) XOR Data[35])));
    OutReady := 1;
    CollectInput(RESET:=TRUE);
  END_IF;
END_PROGRAM

CONFIGURATION Config0
  RESOURCE Res0 ON PLC
    TASK task0(INTERVAL := T#20ms,PRIORITY := 0);
    PROGRAM instance0 WITH task0 : Boiler;
  END_RESOURCE
END_CONFIGURATION

(* ---- RND-EXPR_burgs-hayer-rowan.st ---- *)
(*
This code implements a randomly grown symbolic expression:

((!(!(IN13))) | (!(!(xor(xor(xor(xor(!(IN4 & ((IN19 & true) | (xor(xor(IN42, IN41), IN4)))), xor(xor(!(!(xor(xor(IN31, IN24), IN23))), (xor(xor(xor(xor(IN40, IN28), IN17), IN9), IN39)) & ((IN33 | IN34) & (!(IN20)))), IN44 & ((!(IN32)) & (IN26 & IN44)))), xor(xor(IN11, (IN4 | false) | false), ((xor(xor(IN44, IN24), IN26)) & (!(IN28))) & IN45)), !(xor(xor((xor(xor(IN21, !(IN47)), !(IN8))) | IN40, !(IN1)), xor(xor((IN32 | IN42) & (IN31 & IN45), IN8), xor(xor(false, xor(xor(IN4, IN21), IN1)), !(IN31)))))), xor(xor((!(!(IN26))) | (xor(xor((!(IN37)) | (xor(xor(IN35, IN29), IN14)), (xor(xor(IN20, IN22), IN21)) | (!(IN10))), (!(IN20)) | (IN1 | IN15))), IN15), (((IN24 | IN17) | (xor(xor(IN22, IN33), IN18))) | ((IN15 & IN22) & (IN11 | IN43))) & (!(IN38 | (IN40 & IN44))))))))) & (xor(xor(!((IN45 & (xor(xor(IN43, IN12), true))) & IN23), IN18), xor(xor((((IN22 & (!((IN10 & IN48) & (IN31 & IN35)))) | IN8) & (xor(xor(xor(xor(false, ((IN39 | IN45) | false) & ((IN3 | IN15) & (xor(xor(IN34, IN30), IN33)))), (xor(xor(IN7, IN31 | IN42), IN12 | IN2)) | ((IN4 | IN5) & (IN39 | IN13))), !(IN21 | ((IN20 | IN40) | (IN24 & IN19)))), !(!(xor(xor(IN19, xor(xor(IN37, IN33), IN8)), IN39)))))) | (!(IN35)), !(IN11)), IN45)))

*)

FUNCTION_BLOCK F_CollectInput
  VAR_IN_OUT
      Data : ARRAY[1..50] OF BOOL;
  END_VAR
  VAR_INPUT
      TICK  : BOOL := 0;
      IN1   : BOOL := 0;
      IN2   : BOOL := 0;
      IN3   : BOOL := 0;
      IN4   : BOOL := 0;
      IN5   : BOOL := 0;
      RESET : BOOL := FALSE;
  END_VAR
  VAR_OUTPUT
      Finished : BOOL;
  END_VAR
  VAR
      j    : USINT := 1;
      tock : BOOL  := 0;
  END_VAR
  IF NOT RESET AND tock = NOT TICK THEN
      Data[j]   := IN1;
      Data[j+1] := IN2;
      Data[j+2] := IN3;
      Data[j+3] := IN4;
      Data[j+4] := IN5;
      j := j + 5;
      tock := TICK;
  ELSE
      j := 1;
      tock := 0;
  END_IF;
  Finished := (j > 50);
END_FUNCTION_BLOCK

PROGRAM Boiler
  VAR
    Data  : ARRAY[1..50] OF BOOL;
    Ready : BOOL;
    CollectInput : F_CollectInput;
  END_VAR
  VAR
    TICK     AT %IX1.0 : BOOL;
    IN1      AT %IX0.3 : BOOL;
    IN2      AT %IX0.4 : BOOL;
    IN3      AT %IX0.5 : BOOL;
    IN4      AT %IX0.6 : BOOL;
    IN5      AT %IX0.7 : BOOL;
    OutReady AT %QX0.0 : BOOL := FALSE;
    FeedNext AT %QX0.1 : BOOL := FALSE;
    Out      AT %QX0.2 : BOOL;
  END_VAR
  CollectInput(TICK:=TICK, IN1:=IN1, IN2:=IN2, IN3:=IN3, IN4:=IN4, IN5:=IN5);
  Ready := CollectInput.Finished;
  FeedNext := 1;
  IF Ready THEN
    Out := (((NOT (NOT Data[13])) OR (NOT (NOT (((((NOT (Data[4] AND ((Data[19] AND TRUE) OR ((Data[42] XOR Data[41]) XOR Data[4])))) XOR (((NOT (NOT ((Data[31] XOR Data[24]) XOR Data[23]))) XOR (((((Data[40] XOR Data[28]) XOR Data[17]) XOR Data[9]) XOR Data[39]) AND ((Data[33] OR Data[34]) AND (NOT Data[20])))) XOR (Data[44] AND ((NOT Data[32]) AND (Data[26] AND Data[44]))))) XOR ((Data[11] XOR ((Data[4] OR FALSE) OR FALSE)) XOR ((((Data[44] XOR Data[24]) XOR Data[26]) AND (NOT Data[28])) AND Data[45]))) XOR (NOT (((((Data[21] XOR (NOT Data[47])) XOR (NOT Data[8])) OR Data[40]) XOR (NOT Data[1])) XOR ((((Data[32] OR Data[42]) AND (Data[31] AND Data[45])) XOR Data[8]) XOR ((FALSE XOR ((Data[4] XOR Data[21]) XOR Data[1])) XOR (NOT Data[31])))))) XOR ((((NOT (NOT Data[26])) OR ((((NOT Data[37]) OR ((Data[35] XOR Data[29]) XOR Data[14])) XOR (((Data[20] XOR Data[22]) XOR Data[21]) OR (NOT Data[10]))) XOR ((NOT Data[20]) OR (Data[1] OR Data[15])))) XOR Data[15]) XOR ((((Data[24] OR Data[17]) OR ((Data[22] XOR Data[33]) XOR Data[18])) OR ((Data[15] AND Data[22]) AND (Data[11] OR Data[43]))) AND (NOT (Data[38] OR (Data[40] AND Data[44]))))))))) AND (((NOT ((Data[45] AND ((Data[43] XOR Data[12]) XOR TRUE)) AND Data[23])) XOR Data[18]) XOR ((((((Data[22] AND (NOT ((Data[10] AND Data[48]) AND (Data[31] AND Data[35])))) OR Data[8]) AND ((((FALSE XOR (((Data[39] OR Data[45]) OR FALSE) AND ((Data[3] OR Data[15]) AND ((Data[34] XOR Data[30]) XOR Data[33])))) XOR (((Data[7] XOR (Data[31] OR Data[42])) XOR (Data[12] OR Data[2])) OR ((Data[4] OR Data[5]) AND (Data[39] OR Data[13])))) XOR (NOT (Data[21] OR ((Data[20] OR Data[40]) OR (Data[24] AND Data[19]))))) XOR (NOT (NOT ((Data[19] XOR ((Data[37] XOR Data[33]) XOR Data[8])) XOR Data[39]))))) OR (NOT Data[35])) XOR (NOT Data[11])) XOR Data[45])));
    OutReady := 1;
    CollectInput(RESET:=TRUE);
  END_IF;
END_PROGRAM

CONFIGURATION Config0
  RESOURCE Res0 ON PLC
    TASK task0(INTERVAL := T#20ms,PRIORITY := 0);
    PROGRAM instance0 WITH task0 : Boiler;
  END_RESOURCE
END_CONFIGURATION

(* ---- RND-EXPR_busby-swill-rowed.st ---- *)
(*
This code implements a randomly grown symbolic expression:

(!((!(IN3)) & ((((!(xor(xor(xor(xor(xor(xor(IN22, IN40), IN38), !(IN44)), IN20), IN22), xor(xor(!(IN6), true & IN32), !(IN17))))) | IN31) | (IN3 | IN14)) | IN48))) | ((((!(IN45 & (((xor(xor(IN37 & IN23, IN35), IN11 & IN15)) & IN46) | ((!(IN28 | IN33)) | (!(!(IN13))))))) & IN19) & ((((xor(xor(IN22, !(!(IN40 & IN38))), (xor(xor(IN11 & IN33, IN46 | IN15), IN35 & IN15)) | (!(IN15 | IN17)))) & (!(((IN2 & IN17) | (!(IN16))) & IN16))) & (IN40 | IN25)) & true)) | (xor(xor(IN40, IN11), IN10)))

*)

FUNCTION_BLOCK F_CollectInput
  VAR_IN_OUT
      Data : ARRAY[1..50] OF BOOL;
  END_VAR
  VAR_INPUT
      TICK  : BOOL := 0;
      IN1   : BOOL := 0;
      IN2   : BOOL := 0;
      IN3   : BOOL := 0;
      IN4   : BOOL := 0;
      IN5   : BOOL := 0;
      RESET : BOOL := FALSE;
  END_VAR
  VAR_OUTPUT
      Finished : BOOL;
  END_VAR
  VAR
      j    : USINT := 1;
      tock : BOOL  := 0;
  END_VAR
  IF NOT RESET AND tock = NOT TICK THEN
      Data[j]   := IN1;
      Data[j+1] := IN2;
      Data[j+2] := IN3;
      Data[j+3] := IN4;
      Data[j+4] := IN5;
      j := j + 5;
      tock := TICK;
  ELSE
      j := 1;
      tock := 0;
  END_IF;
  Finished := (j > 50);
END_FUNCTION_BLOCK

PROGRAM Boiler
  VAR
    Data  : ARRAY[1..50] OF BOOL;
    Ready : BOOL;
    CollectInput : F_CollectInput;
  END_VAR
  VAR
    TICK     AT %IX1.0 : BOOL;
    IN1      AT %IX0.3 : BOOL;
    IN2      AT %IX0.4 : BOOL;
    IN3      AT %IX0.5 : BOOL;
    IN4      AT %IX0.6 : BOOL;
    IN5      AT %IX0.7 : BOOL;
    OutReady AT %QX0.0 : BOOL := FALSE;
    FeedNext AT %QX0.1 : BOOL := FALSE;
    Out      AT %QX0.2 : BOOL;
  END_VAR
  CollectInput(TICK:=TICK, IN1:=IN1, IN2:=IN2, IN3:=IN3, IN4:=IN4, IN5:=IN5);
  Ready := CollectInput.Finished;
  FeedNext := 1;
  IF Ready THEN
    Out := ((NOT ((NOT Data[3]) AND ((((NOT ((((((Data[22] XOR Data[40]) XOR Data[38]) XOR (NOT Data[44])) XOR Data[20]) XOR Data[22]) XOR (((NOT Data[6]) XOR (TRUE AND Data[32])) XOR (NOT Data[17])))) OR Data[31]) OR (Data[3] OR Data[14])) OR Data[48]))) OR ((((NOT (Data[45] AND (((((Data[37] AND Data[23]) XOR Data[35]) XOR (Data[11] AND Data[15])) AND Data[46]) OR ((NOT (Data[28] OR Data[33])) OR (NOT (NOT Data[13])))))) AND Data[19]) AND (((((Data[22] XOR (NOT (NOT (Data[40] AND Data[38])))) XOR ((((Data[11] AND Data[33]) XOR (Data[46] OR Data[15])) XOR (Data[35] AND Data[15])) OR (NOT (Data[15] OR Data[17])))) AND (NOT (((Data[2] AND Data[17]) OR (NOT Data[16])) AND Data[16]))) AND (Data[40] OR Data[25])) AND TRUE)) OR ((Data[40] XOR Data[11]) XOR Data[10])));
    OutReady := 1;
    CollectInput(RESET:=TRUE);
  END_IF;
END_PROGRAM

CONFIGURATION Config0
  RESOURCE Res0 ON PLC
    TASK task0(INTERVAL := T#20ms,PRIORITY := 0);
    PROGRAM instance0 WITH task0 : Boiler;
  END_RESOURCE
END_CONFIGURATION

(* ---- RND-EXPR_carne-snook-enjoy.st ---- *)
(*
This code implements a randomly grown symbolic expression:

(xor(xor(((!((((!(IN40)) & ((IN33 | IN34) | IN18)) | (xor(xor((xor(xor(IN25, IN48), IN2)) & (IN15 & IN2), IN50), xor(xor(xor(xor(IN21, IN26), IN45), xor(xor(IN8, IN34), IN32)), IN29 | false)))) | ((xor(xor(IN11, !(IN48 & IN30)), xor(xor(IN43, IN34), IN49 | IN50))) | (!((!(IN42)) & (IN15 & IN15)))))) & ((!(IN7 | ((!(xor(xor(IN2, IN30), IN50))) & ((IN48 | IN25) & (IN49 | IN43))))) | IN15)) & IN6, IN40), IN19 | (!(!((xor(xor(IN8 | IN3, IN37), (xor(xor(xor(xor(IN18, IN45), IN5), IN25 | IN45), !(IN50))) | (IN29 | (!(IN21))))) & ((xor(xor(!(!(IN26)), IN21), (!(IN29)) | (IN43 & IN49))) & (((xor(xor(IN7, IN28), IN29)) | (IN27 | IN22)) | (xor(xor(xor(xor(IN48, IN9), IN42), !(IN43)), xor(xor(IN19, IN42), IN46)))))))))) & (!((xor(xor(!((!((IN24 | (IN2 | IN5)) | (!(!(IN15))))) & ((((IN47 | IN17) | IN39) & (xor(xor(!(IN22), IN26), !(IN24)))) | (!((xor(xor(IN17, IN49), true)) & IN22)))), !(IN31)), xor(xor((!(((IN49 & IN25) & (IN17 | IN5)) | (IN28 | (!(IN32))))) & (!((xor(xor(xor(xor(IN43, IN8), IN8), IN11 | IN14), !(IN6))) & (xor(xor(IN18 & IN5, !(IN50)), IN44)))), (IN46 & IN11) | (IN49 & (xor(xor(!(IN15), !(!(IN30))), !(!(IN42)))))), ((!((!(IN50)) & (IN37 & IN1))) | (xor(xor(IN48, (IN5 & IN15) & IN48), IN42))) | (true & ((xor(xor(IN18 | IN41, !(IN8)), xor(xor(IN46, IN5), IN19))) | IN31))))) | ((!(xor(xor(IN35 & (!(!(IN44 & IN20))), (!((xor(xor(IN4, IN27), IN49)) | (!(IN19)))) | (((!(IN9)) & IN37) & (xor(xor(true | IN45, xor(xor(IN38, IN3), IN32)), IN31)))), !(!((!(IN45)) | (xor(xor(false, IN23), IN22))))))) & IN47)))

*)

FUNCTION_BLOCK F_CollectInput
  VAR_IN_OUT
      Data : ARRAY[1..50] OF BOOL;
  END_VAR
  VAR_INPUT
      TICK  : BOOL := 0;
      IN1   : BOOL := 0;
      IN2   : BOOL := 0;
      IN3   : BOOL := 0;
      IN4   : BOOL := 0;
      IN5   : BOOL := 0;
      RESET : BOOL := FALSE;
  END_VAR
  VAR_OUTPUT
      Finished : BOOL;
  END_VAR
  VAR
      j    : USINT := 1;
      tock : BOOL  := 0;
  END_VAR
  IF NOT RESET AND tock = NOT TICK THEN
      Data[j]   := IN1;
      Data[j+1] := IN2;
      Data[j+2] := IN3;
      Data[j+3] := IN4;
      Data[j+4] := IN5;
      j := j + 5;
      tock := TICK;
  ELSE
      j := 1;
      tock := 0;
  END_IF;
  Finished := (j > 50);
END_FUNCTION_BLOCK

PROGRAM Boiler
  VAR
    Data  : ARRAY[1..50] OF BOOL;
    Ready : BOOL;
    CollectInput : F_CollectInput;
  END_VAR
  VAR
    TICK     AT %IX1.0 : BOOL;
    IN1      AT %IX0.3 : BOOL;
    IN2      AT %IX0.4 : BOOL;
    IN3      AT %IX0.5 : BOOL;
    IN4      AT %IX0.6 : BOOL;
    IN5      AT %IX0.7 : BOOL;
    OutReady AT %QX0.0 : BOOL := FALSE;
    FeedNext AT %QX0.1 : BOOL := FALSE;
    Out      AT %QX0.2 : BOOL;
  END_VAR
  CollectInput(TICK:=TICK, IN1:=IN1, IN2:=IN2, IN3:=IN3, IN4:=IN4, IN5:=IN5);
  Ready := CollectInput.Finished;
  FeedNext := 1;
  IF Ready THEN
    Out := ((((((NOT ((((NOT Data[40]) AND ((Data[33] OR Data[34]) OR Data[18])) OR (((((Data[25] XOR Data[48]) XOR Data[2]) AND (Data[15] AND Data[2])) XOR Data[50]) XOR ((((Data[21] XOR Data[26]) XOR Data[45]) XOR ((Data[8] XOR Data[34]) XOR Data[32])) XOR (Data[29] OR FALSE)))) OR (((Data[11] XOR (NOT (Data[48] AND Data[30]))) XOR ((Data[43] XOR Data[34]) XOR (Data[49] OR Data[50]))) OR (NOT ((NOT Data[42]) AND (Data[15] AND Data[15])))))) AND ((NOT (Data[7] OR ((NOT ((Data[2] XOR Data[30]) XOR Data[50])) AND ((Data[48] OR Data[25]) AND (Data[49] OR Data[43]))))) OR Data[15])) AND Data[6]) XOR Data[40]) XOR (Data[19] OR (NOT (NOT ((((Data[8] OR Data[3]) XOR Data[37]) XOR (((((Data[18] XOR Data[45]) XOR Data[5]) XOR (Data[25] OR Data[45])) XOR (NOT Data[50])) OR (Data[29] OR (NOT Data[21])))) AND ((((NOT (NOT Data[26])) XOR Data[21]) XOR ((NOT Data[29]) OR (Data[43] AND Data[49]))) AND ((((Data[7] XOR Data[28]) XOR Data[29]) OR (Data[27] OR Data[22])) OR ((((Data[48] XOR Data[9]) XOR Data[42]) XOR (NOT Data[43])) XOR ((Data[19] XOR Data[42]) XOR Data[46]))))))))) AND (NOT ((((NOT ((NOT ((Data[24] OR (Data[2] OR Data[5])) OR (NOT (NOT Data[15])))) AND ((((Data[47] OR Data[17]) OR Data[39]) AND (((NOT Data[22]) XOR Data[26]) XOR (NOT Data[24]))) OR (NOT (((Data[17] XOR Data[49]) XOR TRUE) AND Data[22]))))) XOR (NOT Data[31])) XOR ((((NOT (((Data[49] AND Data[25]) AND (Data[17] OR Data[5])) OR (Data[28] OR (NOT Data[32])))) AND (NOT (((((Data[43] XOR Data[8]) XOR Data[8]) XOR (Data[11] OR Data[14])) XOR (NOT Data[6])) AND (((Data[18] AND Data[5]) XOR (NOT Data[50])) XOR Data[44])))) XOR ((Data[46] AND Data[11]) OR (Data[49] AND (((NOT Data[15]) XOR (NOT (NOT Data[30]))) XOR (NOT (NOT Data[42])))))) XOR (((NOT ((NOT Data[50]) AND (Data[37] AND Data[1]))) OR ((Data[48] XOR ((Data[5] AND Data[15]) AND Data[48])) XOR Data[42])) OR (TRUE AND ((((Data[18] OR Data[41]) XOR (NOT Data[8])) XOR ((Data[46] XOR Data[5]) XOR Data[19])) OR Data[31]))))) OR ((NOT (((Data[35] AND (NOT (NOT (Data[44] AND Data[20])))) XOR ((NOT (((Data[4] XOR Data[27]) XOR Data[49]) OR (NOT Data[19]))) OR (((NOT Data[9]) AND Data[37]) AND (((TRUE OR Data[45]) XOR ((Data[38] XOR Data[3]) XOR Data[32])) XOR Data[31])))) XOR (NOT (NOT ((NOT Data[45]) OR ((FALSE XOR Data[23]) XOR Data[22])))))) AND Data[47]))));
    OutReady := 1;
    CollectInput(RESET:=TRUE);
  END_IF;
END_PROGRAM

CONFIGURATION Config0
  RESOURCE Res0 ON PLC
    TASK task0(INTERVAL := T#20ms,PRIORITY := 0);
    PROGRAM instance0 WITH task0 : Boiler;
  END_RESOURCE
END_CONFIGURATION

(* ---- RND-EXPR_casas-obese-clams.st ---- *)
(*
This code implements a randomly grown symbolic expression:

((!(((IN43 | ((xor(xor((IN43 & IN37) & IN9, xor(xor(!(IN43), xor(xor(IN47, IN25), IN19)), !(IN22))), !(IN49 | IN12))) & (IN18 & (!(xor(xor(IN5, IN47), IN46)))))) | (!((((xor(xor(IN17, IN5), IN40)) & true) & IN6) & (!((IN30 & IN17) | (!(IN17))))))) | IN32)) & ((xor(xor((xor(xor((!(xor(xor(IN40, IN40 & IN20), IN30))) & (((IN37 | IN33) | (!(IN46))) & (!(IN7 | IN34))), xor(xor(((IN40 & IN17) | (IN1 | IN24)) & false, IN4), xor(xor((xor(xor(IN3, IN37), IN21)) & (xor(xor(true, IN16), IN32)), (!(IN33)) | (xor(xor(IN45, IN45), IN19))), (IN10 & IN23) | (!(IN37))))), !(xor(xor((IN30 | IN14) | (!(IN15)), (IN8 & IN40) | (IN8 | IN17)), !(xor(xor(IN27, IN47), IN9)))))) | (((!(IN43 | (!(IN37)))) & (!(xor(xor(IN21 | IN17, IN28 & IN4), xor(xor(IN40, IN35), IN2))))) | (!(xor(xor((IN44 | IN34) | IN1, (IN10 | IN32) & IN6), (IN3 & IN35) & (!(IN36)))))), xor(xor(!((xor(xor((IN2 & IN10) | (IN20 & IN9), !(IN15)), IN16)) & IN6), (xor(xor(((!(IN1)) & (IN50 | IN47)) | (IN25 & (!(IN17))), !(IN38)), IN42)) & (((xor(xor(xor(xor(IN2, IN45), true), IN5), !(IN16))) | (!(IN37 & IN5))) | (IN28 & ((xor(xor(IN8, IN33), IN34)) | (xor(xor(IN6, IN3), IN35)))))), !((xor(xor(!(xor(xor(IN2, IN35), IN12)), IN39 & IN15), IN16)) & IN39))), (!(IN11 | ((IN23 & (IN4 | IN3)) | ((IN12 & IN46) & IN3)))) & (!((!(!(IN29 | IN21))) | IN44)))) | (IN33 | (xor(xor((!((xor(xor(IN37 & IN38, xor(xor(IN22, IN46), IN31)), IN41 & IN45)) | (xor(xor(IN26 & IN39, IN46), IN7 | IN38)))) & ((!(!(xor(xor(IN36, IN12), IN27)))) & (!((IN28 & IN23) | (!(IN44))))), IN25), IN49 & (xor(xor(IN38, (xor(xor(IN34, IN30 | IN11), IN6 & IN27)) & (IN18 | (IN16 | IN43))), !((IN30 | IN25) & (xor(xor(IN27, IN31), IN4)))))))))) | (xor(xor(!((!(IN26)) | (!((IN27 & ((!(IN5 | IN16)) & (!(!(IN19))))) | IN21))), IN37), IN21))

*)

FUNCTION_BLOCK F_CollectInput
  VAR_IN_OUT
      Data : ARRAY[1..50] OF BOOL;
  END_VAR
  VAR_INPUT
      TICK  : BOOL := 0;
      IN1   : BOOL := 0;
      IN2   : BOOL := 0;
      IN3   : BOOL := 0;
      IN4   : BOOL := 0;
      IN5   : BOOL := 0;
      RESET : BOOL := FALSE;
  END_VAR
  VAR_OUTPUT
      Finished : BOOL;
  END_VAR
  VAR
      j    : USINT := 1;
      tock : BOOL  := 0;
  END_VAR
  IF NOT RESET AND tock = NOT TICK THEN
      Data[j]   := IN1;
      Data[j+1] := IN2;
      Data[j+2] := IN3;
      Data[j+3] := IN4;
      Data[j+4] := IN5;
      j := j + 5;
      tock := TICK;
  ELSE
      j := 1;
      tock := 0;
  END_IF;
  Finished := (j > 50);
END_FUNCTION_BLOCK

PROGRAM Boiler
  VAR
    Data  : ARRAY[1..50] OF BOOL;
    Ready : BOOL;
    CollectInput : F_CollectInput;
  END_VAR
  VAR
    TICK     AT %IX1.0 : BOOL;
    IN1      AT %IX0.3 : BOOL;
    IN2      AT %IX0.4 : BOOL;
    IN3      AT %IX0.5 : BOOL;
    IN4      AT %IX0.6 : BOOL;
    IN5      AT %IX0.7 : BOOL;
    OutReady AT %QX0.0 : BOOL := FALSE;
    FeedNext AT %QX0.1 : BOOL := FALSE;
    Out      AT %QX0.2 : BOOL;
  END_VAR
  CollectInput(TICK:=TICK, IN1:=IN1, IN2:=IN2, IN3:=IN3, IN4:=IN4, IN5:=IN5);
  Ready := CollectInput.Finished;
  FeedNext := 1;
  IF Ready THEN
    Out := (((NOT (((Data[43] OR (((((Data[43] AND Data[37]) AND Data[9]) XOR (((NOT Data[43]) XOR ((Data[47] XOR Data[25]) XOR Data[19])) XOR (NOT Data[22]))) XOR (NOT (Data[49] OR Data[12]))) AND (Data[18] AND (NOT ((Data[5] XOR Data[47]) XOR Data[46]))))) OR (NOT (((((Data[17] XOR Data[5]) XOR Data[40]) AND TRUE) AND Data[6]) AND (NOT ((Data[30] AND Data[17]) OR (NOT Data[17])))))) OR Data[32])) AND ((((((((NOT ((Data[40] XOR (Data[40] AND Data[20])) XOR Data[30])) AND (((Data[37] OR Data[33]) OR (NOT Data[46])) AND (NOT (Data[7] OR Data[34])))) XOR (((((Data[40] AND Data[17]) OR (Data[1] OR Data[24])) AND FALSE) XOR Data[4]) XOR (((((Data[3] XOR Data[37]) XOR Data[21]) AND ((TRUE XOR Data[16]) XOR Data[32])) XOR ((NOT Data[33]) OR ((Data[45] XOR Data[45]) XOR Data[19]))) XOR ((Data[10] AND Data[23]) OR (NOT Data[37]))))) XOR (NOT ((((Data[30] OR Data[14]) OR (NOT Data[15])) XOR ((Data[8] AND Data[40]) OR (Data[8] OR Data[17]))) XOR (NOT ((Data[27] XOR Data[47]) XOR Data[9]))))) OR (((NOT (Data[43] OR (NOT Data[37]))) AND (NOT (((Data[21] OR Data[17]) XOR (Data[28] AND Data[4])) XOR ((Data[40] XOR Data[35]) XOR Data[2])))) OR (NOT ((((Data[44] OR Data[34]) OR Data[1]) XOR ((Data[10] OR Data[32]) AND Data[6])) XOR ((Data[3] AND Data[35]) AND (NOT Data[36])))))) XOR (((NOT (((((Data[2] AND Data[10]) OR (Data[20] AND Data[9])) XOR (NOT Data[15])) XOR Data[16]) AND Data[6])) XOR ((((((NOT Data[1]) AND (Data[50] OR Data[47])) OR (Data[25] AND (NOT Data[17]))) XOR (NOT Data[38])) XOR Data[42]) AND ((((((Data[2] XOR Data[45]) XOR TRUE) XOR Data[5]) XOR (NOT Data[16])) OR (NOT (Data[37] AND Data[5]))) OR (Data[28] AND (((Data[8] XOR Data[33]) XOR Data[34]) OR ((Data[6] XOR Data[3]) XOR Data[35])))))) XOR (NOT ((((NOT ((Data[2] XOR Data[35]) XOR Data[12])) XOR (Data[39] AND Data[15])) XOR Data[16]) AND Data[39])))) XOR ((NOT (Data[11] OR ((Data[23] AND (Data[4] OR Data[3])) OR ((Data[12] AND Data[46]) AND Data[3])))) AND (NOT ((NOT (NOT (Data[29] OR Data[21]))) OR Data[44])))) OR (Data[33] OR ((((NOT ((((Data[37] AND Data[38]) XOR ((Data[22] XOR Data[46]) XOR Data[31])) XOR (Data[41] AND Data[45])) OR (((Data[26] AND Data[39]) XOR Data[46]) XOR (Data[7] OR Data[38])))) AND ((NOT (NOT ((Data[36] XOR Data[12]) XOR Data[27]))) AND (NOT ((Data[28] AND Data[23]) OR (NOT Data[44]))))) XOR Data[25]) XOR (Data[49] AND ((Data[38] XOR (((Data[34] XOR (Data[30] OR Data[11])) XOR (Data[6] AND Data[27])) AND (Data[18] OR (Data[16] OR Data[43])))) XOR (NOT ((Data[30] OR Data[25]) AND ((Data[27] XOR Data[31]) XOR Data[4]))))))))) OR (((NOT ((NOT Data[26]) OR (NOT ((Data[27] AND ((NOT (Data[5] OR Data[16])) AND (NOT (NOT Data[19])))) OR Data[21])))) XOR Data[37]) XOR Data[21]));
    OutReady := 1;
    CollectInput(RESET:=TRUE);
  END_IF;
END_PROGRAM

CONFIGURATION Config0
  RESOURCE Res0 ON PLC
    TASK task0(INTERVAL := T#20ms,PRIORITY := 0);
    PROGRAM instance0 WITH task0 : Boiler;
  END_RESOURCE
END_CONFIGURATION

(* ---- RND-EXPR_churl-reeky-harsh.st ---- *)
(*
This code implements a randomly grown symbolic expression:

(!(((xor(xor((!(xor(xor((!(IN37)) | (xor(xor(IN14, IN5), IN24)), (IN12 & IN29) | (IN14 & IN43)), (IN49 | IN19) & IN19))) | (!(((!(IN6)) | (IN47 & IN17)) | ((xor(xor(IN7, IN8), IN40)) | IN39))), (xor(xor(xor(xor(xor(xor(!(IN50), IN18), xor(xor(IN23, IN45), IN35)), (IN20 | IN15) & IN30), IN32), ((IN8 | IN22) & (IN32 | IN18)) & (!(IN9 | IN37))), xor(xor(!(true & IN23), IN42 | (!(IN49))), xor(xor(xor(xor(IN25, IN20), IN2), !(IN29)), IN35 | IN42)))) & IN31), !(!((IN12 | (IN45 & IN17)) & ((IN32 & IN23) | (IN3 & IN27)))))) & (!((xor(xor(true, ((IN26 & IN1) | (!(IN34))) & IN44), !(IN22))) | (!(IN38))))) & ((!(!(xor(xor(IN39 & ((xor(xor(IN26, IN47), IN31)) & (IN15 | IN46)), !((IN44 & IN5) & IN31)), IN30)))) & (!((xor(xor(!((IN39 & IN2) & (xor(xor(IN15, IN17), IN26))), !(IN47)), ((!(IN31)) | (!(IN38))) & (xor(xor(IN45 & IN39, xor(xor(IN33, IN15), IN16)), xor(xor(IN34, IN46), IN20))))) & (((xor(xor(IN48 & IN33, !(IN44)), IN34)) | IN29) | ((xor(xor(!(IN1), IN47 | IN15), IN4 | IN9)) | IN37))))))) | IN5

*)

FUNCTION_BLOCK F_CollectInput
  VAR_IN_OUT
      Data : ARRAY[1..50] OF BOOL;
  END_VAR
  VAR_INPUT
      TICK  : BOOL := 0;
      IN1   : BOOL := 0;
      IN2   : BOOL := 0;
      IN3   : BOOL := 0;
      IN4   : BOOL := 0;
      IN5   : BOOL := 0;
      RESET : BOOL := FALSE;
  END_VAR
  VAR_OUTPUT
      Finished : BOOL;
  END_VAR
  VAR
      j    : USINT := 1;
      tock : BOOL  := 0;
  END_VAR
  IF NOT RESET AND tock = NOT TICK THEN
      Data[j]   := IN1;
      Data[j+1] := IN2;
      Data[j+2] := IN3;
      Data[j+3] := IN4;
      Data[j+4] := IN5;
      j := j + 5;
      tock := TICK;
  ELSE
      j := 1;
      tock := 0;
  END_IF;
  Finished := (j > 50);
END_FUNCTION_BLOCK

PROGRAM Boiler
  VAR
    Data  : ARRAY[1..50] OF BOOL;
    Ready : BOOL;
    CollectInput : F_CollectInput;
  END_VAR
  VAR
    TICK     AT %IX1.0 : BOOL;
    IN1      AT %IX0.3 : BOOL;
    IN2      AT %IX0.4 : BOOL;
    IN3      AT %IX0.5 : BOOL;
    IN4      AT %IX0.6 : BOOL;
    IN5      AT %IX0.7 : BOOL;
    OutReady AT %QX0.0 : BOOL := FALSE;
    FeedNext AT %QX0.1 : BOOL := FALSE;
    Out      AT %QX0.2 : BOOL;
  END_VAR
  CollectInput(TICK:=TICK, IN1:=IN1, IN2:=IN2, IN3:=IN3, IN4:=IN4, IN5:=IN5);
  Ready := CollectInput.Finished;
  FeedNext := 1;
  IF Ready THEN
    Out := ((NOT ((((((NOT ((((NOT Data[37]) OR ((Data[14] XOR Data[5]) XOR Data[24])) XOR ((Data[12] AND Data[29]) OR (Data[14] AND Data[43]))) XOR ((Data[49] OR Data[19]) AND Data[19]))) OR (NOT (((NOT Data[6]) OR (Data[47] AND Data[17])) OR (((Data[7] XOR Data[8]) XOR Data[40]) OR Data[39])))) XOR ((((((((NOT Data[50]) XOR Data[18]) XOR ((Data[23] XOR Data[45]) XOR Data[35])) XOR ((Data[20] OR Data[15]) AND Data[30])) XOR Data[32]) XOR (((Data[8] OR Data[22]) AND (Data[32] OR Data[18])) AND (NOT (Data[9] OR Data[37])))) XOR (((NOT (TRUE AND Data[23])) XOR (Data[42] OR (NOT Data[49]))) XOR ((((Data[25] XOR Data[20]) XOR Data[2]) XOR (NOT Data[29])) XOR (Data[35] OR Data[42])))) AND Data[31])) XOR (NOT (NOT ((Data[12] OR (Data[45] AND Data[17])) AND ((Data[32] AND Data[23]) OR (Data[3] AND Data[27])))))) AND (NOT (((TRUE XOR (((Data[26] AND Data[1]) OR (NOT Data[34])) AND Data[44])) XOR (NOT Data[22])) OR (NOT Data[38])))) AND ((NOT (NOT (((Data[39] AND (((Data[26] XOR Data[47]) XOR Data[31]) AND (Data[15] OR Data[46]))) XOR (NOT ((Data[44] AND Data[5]) AND Data[31]))) XOR Data[30]))) AND (NOT ((((NOT ((Data[39] AND Data[2]) AND ((Data[15] XOR Data[17]) XOR Data[26]))) XOR (NOT Data[47])) XOR (((NOT Data[31]) OR (NOT Data[38])) AND (((Data[45] AND Data[39]) XOR ((Data[33] XOR Data[15]) XOR Data[16])) XOR ((Data[34] XOR Data[46]) XOR Data[20])))) AND (((((Data[48] AND Data[33]) XOR (NOT Data[44])) XOR Data[34]) OR Data[29]) OR ((((NOT Data[1]) XOR (Data[47] OR Data[15])) XOR (Data[4] OR Data[9])) OR Data[37]))))))) OR Data[5]);
    OutReady := 1;
    CollectInput(RESET:=TRUE);
  END_IF;
END_PROGRAM

CONFIGURATION Config0
  RESOURCE Res0 ON PLC
    TASK task0(INTERVAL := T#20ms,PRIORITY := 0);
    PROGRAM instance0 WITH task0 : Boiler;
  END_RESOURCE
END_CONFIGURATION

(* ---- RND-EXPR_clerk-chump-agile.st ---- *)
(*
This code implements a randomly grown symbolic expression:

IN42 | (xor(xor(!((xor(xor((((xor(xor(IN16, IN3 | IN21), IN3 & IN18)) & ((IN42 & IN40) & (xor(xor(IN43, IN4), IN7)))) | (!((IN49 | IN47) | (xor(xor(IN2, IN11), IN5))))) | (xor(xor(!((true & IN23) & (IN45 | IN1)), IN13 & ((!(IN21)) & (IN48 & IN18))), ((xor(xor(IN21, IN4), IN7)) | (!(IN40))) & ((IN3 | IN27) | (IN16 | IN44)))), IN9), IN3)) & IN50), IN19), IN13))

*)

FUNCTION_BLOCK F_CollectInput
  VAR_IN_OUT
      Data : ARRAY[1..50] OF BOOL;
  END_VAR
  VAR_INPUT
      TICK  : BOOL := 0;
      IN1   : BOOL := 0;
      IN2   : BOOL := 0;
      IN3   : BOOL := 0;
      IN4   : BOOL := 0;
      IN5   : BOOL := 0;
      RESET : BOOL := FALSE;
  END_VAR
  VAR_OUTPUT
      Finished : BOOL;
  END_VAR
  VAR
      j    : USINT := 1;
      tock : BOOL  := 0;
  END_VAR
  IF NOT RESET AND tock = NOT TICK THEN
      Data[j]   := IN1;
      Data[j+1] := IN2;
      Data[j+2] := IN3;
      Data[j+3] := IN4;
      Data[j+4] := IN5;
      j := j + 5;
      tock := TICK;
  ELSE
      j := 1;
      tock := 0;
  END_IF;
  Finished := (j > 50);
END_FUNCTION_BLOCK

PROGRAM Boiler
  VAR
    Data  : ARRAY[1..50] OF BOOL;
    Ready : BOOL;
    CollectInput : F_CollectInput;
  END_VAR
  VAR
    TICK     AT %IX1.0 : BOOL;
    IN1      AT %IX0.3 : BOOL;
    IN2      AT %IX0.4 : BOOL;
    IN3      AT %IX0.5 : BOOL;
    IN4      AT %IX0.6 : BOOL;
    IN5      AT %IX0.7 : BOOL;
    OutReady AT %QX0.0 : BOOL := FALSE;
    FeedNext AT %QX0.1 : BOOL := FALSE;
    Out      AT %QX0.2 : BOOL;
  END_VAR
  CollectInput(TICK:=TICK, IN1:=IN1, IN2:=IN2, IN3:=IN3, IN4:=IN4, IN5:=IN5);
  Ready := CollectInput.Finished;
  FeedNext := 1;
  IF Ready THEN
    Out := (Data[42] OR (((NOT ((((((((Data[16] XOR (Data[3] OR Data[21])) XOR (Data[3] AND Data[18])) AND ((Data[42] AND Data[40]) AND ((Data[43] XOR Data[4]) XOR Data[7]))) OR (NOT ((Data[49] OR Data[47]) OR ((Data[2] XOR Data[11]) XOR Data[5])))) OR (((NOT ((TRUE AND Data[23]) AND (Data[45] OR Data[1]))) XOR (Data[13] AND ((NOT Data[21]) AND (Data[48] AND Data[18])))) XOR ((((Data[21] XOR Data[4]) XOR Data[7]) OR (NOT Data[40])) AND ((Data[3] OR Data[27]) OR (Data[16] OR Data[44]))))) XOR Data[9]) XOR Data[3]) AND Data[50])) XOR Data[19]) XOR Data[13]));
    OutReady := 1;
    CollectInput(RESET:=TRUE);
  END_IF;
END_PROGRAM

CONFIGURATION Config0
  RESOURCE Res0 ON PLC
    TASK task0(INTERVAL := T#20ms,PRIORITY := 0);
    PROGRAM instance0 WITH task0 : Boiler;
  END_RESOURCE
END_CONFIGURATION

(* ---- RND-EXPR_click-grief-pubis.st ---- *)
(*
This code implements a randomly grown symbolic expression:

(xor(xor(IN40, IN23), IN33)) | IN36

*)

FUNCTION_BLOCK F_CollectInput
  VAR_IN_OUT
      Data : ARRAY[1..50] OF BOOL;
  END_VAR
  VAR_INPUT
      TICK  : BOOL := 0;
      IN1   : BOOL := 0;
      IN2   : BOOL := 0;
      IN3   : BOOL := 0;
      IN4   : BOOL := 0;
      IN5   : BOOL := 0;
      RESET : BOOL := FALSE;
  END_VAR
  VAR_OUTPUT
      Finished : BOOL;
  END_VAR
  VAR
      j    : USINT := 1;
      tock : BOOL  := 0;
  END_VAR
  IF NOT RESET AND tock = NOT TICK THEN
      Data[j]   := IN1;
      Data[j+1] := IN2;
      Data[j+2] := IN3;
      Data[j+3] := IN4;
      Data[j+4] := IN5;
      j := j + 5;
      tock := TICK;
  ELSE
      j := 1;
      tock := 0;
  END_IF;
  Finished := (j > 50);
END_FUNCTION_BLOCK

PROGRAM Boiler
  VAR
    Data  : ARRAY[1..50] OF BOOL;
    Ready : BOOL;
    CollectInput : F_CollectInput;
  END_VAR
  VAR
    TICK     AT %IX1.0 : BOOL;
    IN1      AT %IX0.3 : BOOL;
    IN2      AT %IX0.4 : BOOL;
    IN3      AT %IX0.5 : BOOL;
    IN4      AT %IX0.6 : BOOL;
    IN5      AT %IX0.7 : BOOL;
    OutReady AT %QX0.0 : BOOL := FALSE;
    FeedNext AT %QX0.1 : BOOL := FALSE;
    Out      AT %QX0.2 : BOOL;
  END_VAR
  CollectInput(TICK:=TICK, IN1:=IN1, IN2:=IN2, IN3:=IN3, IN4:=IN4, IN5:=IN5);
  Ready := CollectInput.Finished;
  FeedNext := 1;
  IF Ready THEN
    Out := (((Data[40] XOR Data[23]) XOR Data[33]) OR Data[36]);
    OutReady := 1;
    CollectInput(RESET:=TRUE);
  END_IF;
END_PROGRAM

CONFIGURATION Config0
  RESOURCE Res0 ON PLC
    TASK task0(INTERVAL := T#20ms,PRIORITY := 0);
    PROGRAM instance0 WITH task0 : Boiler;
  END_RESOURCE
END_CONFIGURATION

(* ---- RND-EXPR_coper-ravel-devil.st ---- *)
(*
This code implements a randomly grown symbolic expression:

!(IN17)

*)

FUNCTION_BLOCK F_CollectInput
  VAR_IN_OUT
      Data : ARRAY[1..50] OF BOOL;
  END_VAR
  VAR_INPUT
      TICK  : BOOL := 0;
      IN1   : BOOL := 0;
      IN2   : BOOL := 0;
      IN3   : BOOL := 0;
      IN4   : BOOL := 0;
      IN5   : BOOL := 0;
      RESET : BOOL := FALSE;
  END_VAR
  VAR_OUTPUT
      Finished : BOOL;
  END_VAR
  VAR
      j    : USINT := 1;
      tock : BOOL  := 0;
  END_VAR
  IF NOT RESET AND tock = NOT TICK THEN
      Data[j]   := IN1;
      Data[j+1] := IN2;
      Data[j+2] := IN3;
      Data[j+3] := IN4;
      Data[j+4] := IN5;
      j := j + 5;
      tock := TICK;
  ELSE
      j := 1;
      tock := 0;
  END_IF;
  Finished := (j > 50);
END_FUNCTION_BLOCK

PROGRAM Boiler
  VAR
    Data  : ARRAY[1..50] OF BOOL;
    Ready : BOOL;
    CollectInput : F_CollectInput;
  END_VAR
  VAR
    TICK     AT %IX1.0 : BOOL;
    IN1      AT %IX0.3 : BOOL;
    IN2      AT %IX0.4 : BOOL;
    IN3      AT %IX0.5 : BOOL;
    IN4      AT %IX0.6 : BOOL;
    IN5      AT %IX0.7 : BOOL;
    OutReady AT %QX0.0 : BOOL := FALSE;
    FeedNext AT %QX0.1 : BOOL := FALSE;
    Out      AT %QX0.2 : BOOL;
  END_VAR
  CollectInput(TICK:=TICK, IN1:=IN1, IN2:=IN2, IN3:=IN3, IN4:=IN4, IN5:=IN5);
  Ready := CollectInput.Finished;
  FeedNext := 1;
  IF Ready THEN
    Out := (NOT Data[17]);
    OutReady := 1;
    CollectInput(RESET:=TRUE);
  END_IF;
END_PROGRAM

CONFIGURATION Config0
  RESOURCE Res0 ON PLC
    TASK task0(INTERVAL := T#20ms,PRIORITY := 0);
    PROGRAM instance0 WITH task0 : Boiler;
  END_RESOURCE
END_CONFIGURATION

(* ---- RND-EXPR_count-toils-budge.st ---- *)
(*
This code implements a randomly grown symbolic expression:

!(IN40)

*)

FUNCTION_BLOCK F_CollectInput
  VAR_IN_OUT
      Data : ARRAY[1..50] OF BOOL;
  END_VAR
  VAR_INPUT
      TICK  : BOOL := 0;
      IN1   : BOOL := 0;
      IN2   : BOOL := 0;
      IN3   : BOOL := 0;
      IN4   : BOOL := 0;
      IN5   : BOOL := 0;
      RESET : BOOL := FALSE;
  END_VAR
  VAR_OUTPUT
      Finished : BOOL;
  END_VAR
  VAR
      j    : USINT := 1;
      tock : BOOL  := 0;
  END_VAR
  IF NOT RESET AND tock = NOT TICK THEN
      Data[j]   := IN1;
      Data[j+1] := IN2;
      Data[j+2] := IN3;
      Data[j+3] := IN4;
      Data[j+4] := IN5;
      j := j + 5;
      tock := TICK;
  ELSE
      j := 1;
      tock := 0;
  END_IF;
  Finished := (j > 50);
END_FUNCTION_BLOCK

PROGRAM Boiler
  VAR
    Data  : ARRAY[1..50] OF BOOL;
    Ready : BOOL;
    CollectInput : F_CollectInput;
  END_VAR
  VAR
    TICK     AT %IX1.0 : BOOL;
    IN1      AT %IX0.3 : BOOL;
    IN2      AT %IX0.4 : BOOL;
    IN3      AT %IX0.5 : BOOL;
    IN4      AT %IX0.6 : BOOL;
    IN5      AT %IX0.7 : BOOL;
    OutReady AT %QX0.0 : BOOL := FALSE;
    FeedNext AT %QX0.1 : BOOL := FALSE;
    Out      AT %QX0.2 : BOOL;
  END_VAR
  CollectInput(TICK:=TICK, IN1:=IN1, IN2:=IN2, IN3:=IN3, IN4:=IN4, IN5:=IN5);
  Ready := CollectInput.Finished;
  FeedNext := 1;
  IF Ready THEN
    Out := (NOT Data[40]);
    OutReady := 1;
    CollectInput(RESET:=TRUE);
  END_IF;
END_PROGRAM

CONFIGURATION Config0
  RESOURCE Res0 ON PLC
    TASK task0(INTERVAL := T#20ms,PRIORITY := 0);
    PROGRAM instance0 WITH task0 : Boiler;
  END_RESOURCE
END_CONFIGURATION
